(* IEC 61131-3 sources: daoli-st-library/DL_Process (part 28) *)

(* ---- FB_DL_ChillerYearWinStart.st ---- *)
(*==============================================================================
 * 组件名称 (Component)  : FB_DL_ChillerYearWinStart
 * 所属子库 (Sublibrary) : DL_Process
 * 当前版本 (Version)    : 1.0.0
 * 兼容性 (Platform)     : CODESYS 3.5+ / TwinCAT 3 / 汇川 InoProShop / 施耐德 Machine Expert
 *                         仅依赖 Standard.library（R_TRIG），零厂商私有库
 * 功能描述 (Function)   : 冷机年度启停窗与保养互锁。启动申请仅在「年窗电平
 *                         内 + 保养完成互锁成立」时放行 bRun，否则拒绝并按
 *                         独立成因（非窗 / 保养未完）给出 bBlocked 电平与
 *                         eBlock 成因（R190 归因唯一）；运行中可随时停止。
 *                         与 YearWindowCheck（年窗原子）分工：本件叠加
 *                         「非窗禁启」的设备控制语义。
 * 来源标签 (Origin)     : ROADMAP §16.5 R11 池（L725），自研 clean-room
 * 边界语义 (Boundary)   : ① 启动判据全组合闸（窗电平 / 保养互锁 / 无故障），
 *                         拒启不锁存故障（拒绝是正常业务态）；
 *                         ② 保养互锁输入非有限无涉（布尔域），无浮点量；
 *                         ③ eBlock 成因独立成员逐拍重算（拒绝成因随当前
 *                         条件实时回放，信息级允许每拍重算，R189）。
 * 输出语义 (Fallback)   : 【R191】bEnable = FALSE → bRun 强制 FALSE（启停
 *                         出口失能必须收敛）；eFault 相 → bRun FALSE + bError。
 * 码位     (Codes)      : 按 R297 范式零 16# 码位硬编码；错误出口 BOOL+ENUM(eCause)。
 * 红线自检 (Redline)    : 7 项红线已自检：R1 零全局 ✓｜R2 零物理地址 ✓｜R3 纯 IEC ✓
 *                         R4 无浮点域/组态无涉 ✓｜R5 双语同行注释 ✓
 *                         R6 CASE 带 ELSE 兜底迁 eFault ✓｜R7 R_TRIG 段 0 无条件刷新 ✓
 * 验收向量 (Acceptance) : V1 窗内 + 保养完 + 申请沿 → bRun=TRUE，bBlocked=FALSE；
 *                         V2 窗外申请沿 → bRun=FALSE，bBlocked=TRUE，
 *                         eBlock=eNotInWin；
 *                         V3 窗内但保养未完 → eBlock=eMaintDue（非窗成因
 *                         不再误报）。
 * 修订历史 (Revision)   : 2026-11-20  v1.0.0  R51 首版（批 2 · 序号 7）
 *==============================================================================*)
TYPE E_DL_CwsBlock :
(
    eNone     := 0,                          (* 无拒绝（已放行或无申请） / No block *)
    eNotInWin := 1,                          (* 非年窗禁启 / Not in year window *)
    eMaintDue := 2                           (* 保养未完禁启 / Maintenance interlock open *)
);
END_TYPE

TYPE E_DL_CwsState :
(
    eIdle  := 0,                             (* 停机待窗 / Idle *)
    eRun   := 10,                            (* 运行 / Running *)
    eFault := 90                             (* 故障锁存相 / Fault latched phase *)
);
END_TYPE

TYPE E_DL_CwsCause :
(
    eNone     := 0,                          (* 无故障成因 / No cause *)
    ePhaseBad := 3                           (* 非法相位兜底 / Illegal phase fallback *)
);
END_TYPE

FUNCTION_BLOCK FB_DL_ChillerYearWinStart
VAR_INPUT
    bInWin     : BOOL := FALSE;              (* 年窗电平（上层 YearWindowCheck 供给）[-] / Year-window level *)
    bMaintOk   : BOOL := TRUE;               (* 保养完成互锁电平 [-] / Maintenance interlock *)
    bStartReq  : BOOL := FALSE;              (* 启动申请电平 [-] / Start request *)
    bStopReq   : BOOL := FALSE;              (* 停止申请电平（运行中随时可停）[-] / Stop request *)
    bEnable    : BOOL := TRUE;               (* 使能 [-] / Enable *)
    bReset     : BOOL := FALSE;              (* 复位命令，上升沿清全部 [-] / Reset command *)
END_VAR
VAR_OUTPUT
    bRun       : BOOL;                       (* 冷机运行出口 [-] / Run outlet *)
    bStartOk   : BOOL;                       (* 本次申请放行单拍位 [-] / Start-allowed pulse *)
    bBlocked   : BOOL;                       (* 申请被拒电平（申请期实时）[-] / Blocked level *)
    eBlock     : E_DL_CwsBlock;              (* 拒绝成因（信息级逐拍重算，R189） / Block cause *)
    nRunCycles : UDINT;                      (* 累计启动次数 [次] / Run cycle count *)
    eState     : E_DL_CwsState;              (* 状态出口 / State outlet *)
    eCause     : E_DL_CwsCause;              (* 故障成因出口 / Fault cause outlet *)
    bError     : BOOL;                       (* 故障锁存标志 [-] / Fault latch flag *)
END_VAR
VAR
    _eState   : E_DL_CwsState := E_DL_CwsState.eIdle;     (* 内部相位（CASE 唯一写入目标） / Internal phase *)
    _eCause   : E_DL_CwsCause := E_DL_CwsCause.eNone;     (* 故障成因锁存量 / Latched cause *)
    rtStart   : R_TRIG;                      (* 启动申请沿实例，段 0 无条件调用 / Start edge instance *)
    rtStop    : R_TRIG;                      (* 停止申请沿实例，段 0 无条件调用 / Stop edge instance *)
    rtReset   : R_TRIG;                      (* 复位沿实例，段 0 无条件调用 / Reset edge instance *)
    _nCycles  : UDINT;                       (* 启动计数锁存 [次] / Cycle count latch *)
    _bStartOk : BOOL;                        (* 放行单拍量 [-] / Start-allowed work *)
    _bFault   : BOOL;                        (* 故障锁存位 / Latched fault bit *)
END_VAR

(* —— 段 0：沿实例无条件刷新（R228A；纯布尔域无浮点组态闸） —— *)
rtStart(CLK := bStartReq);                   (* 启动沿每拍必调 / Start edge every scan *)
rtStop(CLK := bStopReq);                     (* 停止沿每拍必调 / Stop edge every scan *)
rtReset(CLK := bReset);                      (* 复位沿每拍必调 / Reset edge every scan *)

(* —— 段 1：单拍量预清零（R107） —— *)
_bStartOk := FALSE;                          (* 放行脉冲预清，唯一分支置位 / Start-ok preset *)
bStartOk := FALSE;                           (* 放行出口预清 / Start-ok outlet preset *)
bBlocked := FALSE;                           (* 拒绝电平预清 / Blocked preset *)
eBlock := E_DL_CwsBlock.eNone;               (* 拒绝成因预清（判定分支覆盖） / Block cause preset *)

(* —— 段 2：复位沿处理（作用域：清故障 + 清计数 + 迁 eIdle（bRun 随相位收敛），R283 逐项声明） —— *)
IF rtReset.Q THEN
    _bFault := FALSE;                        (* 清故障锁存 / Clear fault *)
    _eCause := E_DL_CwsCause.eNone;          (* 清成因 / Clear cause *)
    _nCycles := 0;                           (* 清启动计数 / Clear count *)
    _eState := E_DL_CwsState.eIdle;          (* 迁停机相 / Back to idle *)
END_IF

(* —— 段 4：CASE 主状态机（ELSE 兜底迁 eFault，红线 6） —— *)
CASE _eState OF
    E_DL_CwsState.eIdle:                     (* 停机相 / Idle *)
        IF rtStart.Q AND bEnable THEN        (* 申请沿：判组合闸 / On start edge *)
            IF NOT bInWin THEN
                bBlocked := TRUE;            (* 拒绝电平 / Blocked level *)
                eBlock := E_DL_CwsBlock.eNotInWin;   (* 成因：非窗（独立成员，R190） / Cause: not in window *)
            ELSIF NOT bMaintOk THEN
                bBlocked := TRUE;            (* 拒绝电平 / Blocked level *)
                eBlock := E_DL_CwsBlock.eMaintDue;   (* 成因：保养未完 / Cause: maintenance *)
            ELSE
                _bStartOk := TRUE;           (* 放行单拍 / Start-ok pulse *)
                _nCycles := _nCycles + 1;    (* 启动计数（UDINT 回绕工程安全） / Count start *)
                _eState := E_DL_CwsState.eRun;   (* 进入运行 / Enter run *)
            END_IF
        END_IF
    E_DL_CwsState.eRun:                      (* 运行相：停止沿随时出 / Run *)
        IF rtStop.Q OR (NOT bEnable) THEN    (* 停止沿或失能：回停机 / Stop or disable *)
            _eState := E_DL_CwsState.eIdle;  (* 回停机相 / Back to idle *)
        END_IF
    E_DL_CwsState.eFault:                    (* 故障相：仅复位沿出（bRun 随段 5 收敛） / Fault *)
        ;                                    (* 锁存回放（R28） / Replay from latch *)
    ELSE                                     (* 非法相位兜底迁安全态 / Illegal phase fallback *)
        _eState := E_DL_CwsState.eFault;     (* 迁故障相 / To fault *)
        _bFault := TRUE;                     (* 同步锁存 / Latch *)
        _eCause := E_DL_CwsCause.ePhaseBad;  (* 成因：非法相位 / Cause: illegal phase *)
END_CASE

(* —— 段 5：出口映射（bRun 与相位同源同义，R191 名实双出口） —— *)
bRun := (_eState = E_DL_CwsState.eRun) AND bEnable AND (NOT _bFault);   (* 运行出口（失能/故障收敛 FALSE） / Run outlet *)
bStartOk := _bStartOk;                       (* 放行脉冲出口 / Start-ok outlet *)
nRunCycles := _nCycles;                      (* 启动计数出口 / Count outlet *)
bError := _bFault;                           (* 故障标志镜像 / Fault flag mirror *)
eState := _eState;                           (* 状态出口 / State outlet *)
eCause := _eCause;                           (* 成因出口 / Cause outlet *)
END_FUNCTION_BLOCK

(* ---- FB_DL_CleanRoomPressure.st ---- *)
(*==============================================================================
 * 组件名称 (Component)  : FB_DL_CleanRoomPressure
 * 所属子库 (Sublibrary) : DL_Process
 * 前缀     (Prefix)     : FB_DL_
 * 当前版本 (Version)    : 1.0.0
 * 兼容性   (Platform)   : CODESYS 3.5 / TwinCAT 3 / 汇川 InoProShop / Schneider
 *                         Machine Expert；纯 IEC 61131-3（第 3 版），
 *                         仅依赖标准库 MAX / MIN，零厂商方言、零定时器依赖
 * 作者     (Author)     : 道莅代码库 · PLC编程专家（R31）
 * 开源溯源 (Origin)     : 洁净室压差梯级控制公开工艺语义（行业池），道莅
 *                         clean-room 防御性实现，未复制任何外部源码行
 * 功能描述 (Function)   : 多房间正压梯级控制防倒流件。梯度校验先于控制：
 *                         逐室核对设定梯度沿洁净度递减方向严格递减，
 *                         倒置即锁存倒置标志并冻结投切（防倒流最高优先）；
 *                         控制层各室独立带回差双限：低于下限请求加大风量、
 *                         高于上限撤回请求、带内保持。
 * 码位     (Codes)      : 16#0005_00A3 信息级：压差/设定非有限该室退出仲裁、
 *                                      房间计数钳位（不置 bError）
 *                         16#0005_00A4 故障级：梯度倒置（锁存，独立复位通道）
 *                         16#0005_00A5~00A7 保留未启用（码表与实现对齐）
 * 边界防错 (Boundary)   : 1 梯度倒置锁存有可达解除式：独立 bRstInv 复位沿，
 *                           复位通道不受 NOT bEn 屏蔽（终审两式之一）；
 *                         2 房间计数钳上限、越界逐位清零；
 *                         3 非有限压差该室退出仲裁保持原投切并计掩码；
 *                         4 首拍全 FALSE；
 *                         5 无定时器/边沿实例（纯组合投切层）。
 * 修订历史 (Revision)   : 2026-11-18 v1.0.0 首版入库（R31 · 阶段三 · 序 13）
 *==============================================================================*)

(*==============================================================================
 * 功能块: FB_DL_CleanRoomPressure
 * 调用约定: 每个扫描周期无条件调用一次；压差与梯度设定经引脚数组注入，
 *           数组维度 1..8（8 室上限），有效室数经 uRoomCnt 给出。
 *==============================================================================*)
FUNCTION_BLOCK FB_DL_CleanRoomPressure
VAR_INPUT
    afDp    : ARRAY[1..8] OF REAL;    // 各室实测压差 [帕] / Per-room measured differential pressure [Pa]
    afSet   : ARRAY[1..8] OF REAL;    // 各室压差梯度设定 [帕]，须严格递减 / Per-room gradient setpoints [Pa], strictly decreasing
    uRoomCnt: UINT := 8;              // 有效房间数 [间]，合法域 1..8 / Valid room count, valid 1..8
    fBand   : REAL := 5.0;            // 回差半带宽 [帕] / Hysteresis half band [Pa]
    bEn     : BOOL := FALSE;          // 使能 / Enable flag
    bRstInv : BOOL := FALSE;          // 梯度倒置独立复位沿（不受使能屏蔽）/ Inversion reset edge, never masked by enable
END_VAR
VAR_OUTPUT
    abBoost : ARRAY[1..8] OF BOOL;    // 各室加大风量请求 / Per-room boost request
    bInvert : BOOL;                   // 梯度倒置锁存标志 / Gradient inversion latch flag
    uErrorId: UDINT;                  // 错误码，0 = 无错 / Error code, 0 = none
END_VAR
VAR
    rTrigRst: R_TRIG;                 // 倒置复位沿检测，每拍无条件刷新 / Inversion reset edge detector
    uCntEff : INT;                    // 钳位后有效室数 [间]，INT 域循环 / Effective clamped room count, INT domain
    i       : INT;                    // 逐室循环索引 / Per-room loop index
    bRoomOk : ARRAY[1..8] OF BOOL;    // 各室数据有效掩码 / Per-room data validity mask
    bBadAny : BOOL;                   // 任一室数据无效 / Any room data invalid
    bFirst  : BOOL := TRUE;           // 首拍标志 / First-scan flag
    fLo     : REAL;                   // 本室投切下限 [帕] / Room switching lower bound [Pa]
    fHi     : REAL;                   // 本室投切上限 [帕] / Room switching upper bound [Pa]
END_VAR
VAR CONSTANT
    DL_CRP_ROOM_MAX: INT  := 8;       // 房间数上限 [间] / Room count upper bound
    DL_CRP_FIN     : REAL := 1.0E30;  // REAL 有限幅值判界 / REAL finiteness magnitude bound
END_VAR

// ---- 段 1｜边沿实例无条件刷新（红线：禁入条件分支）----------------------------
rTrigRst(CLK := bRstInv);                             // 倒置复位沿检测 / Inversion reset edge detection

// ---- 段 2｜梯度倒置独立复位：先于一切使能门控（R38 复位通道不屏蔽）--------------
IF rTrigRst.Q THEN
    bInvert := FALSE;                                 // 复位清倒置锁存 / Reset clears inversion latch
END_IF

// ---- 段 3｜计数钳位与首拍初始化 --------------------------------------------------
uCntEff := MIN(UINT_TO_INT(uRoomCnt), DL_CRP_ROOM_MAX); // 计数钳上限，统一 INT 域 / Clamp count, unified INT domain
uCntEff := MAX(uCntEff, 1);                           // 下限保 1 防 0 循环 / Floor at 1 against empty loop
IF bFirst THEN
    FOR i := 1 TO DL_CRP_ROOM_MAX DO
        abBoost[i] := FALSE;                          // 首拍全 FALSE / First scan all FALSE
        bRoomOk[i] := TRUE;                           // 掩码预置有效 / Mask preset valid
    END_FOR
    bFirst := FALSE;                                  // 清首拍标志 / Clear first-scan flag
END_IF

// ---- 段 4｜梯度校验先于控制（防倒流最高优先）--------------------------------------
IF NOT bInvert THEN
    FOR i := 1 TO (uCntEff - 1) DO
        IF (afSet[i] <> afSet[i]) OR (afSet[i + 1] <> afSet[i + 1])
           OR (ABS(afSet[i]) >= DL_CRP_FIN) OR (ABS(afSet[i + 1]) >= DL_CRP_FIN) THEN
            bInvert := TRUE;                          // 非有限设定按倒置保守处理（留档）/ Non-finite set treated as inversion
        ELSIF afSet[i] <= afSet[i + 1] THEN
            bInvert := TRUE;                          // 梯度未严格递减判倒置 / Non-decreasing gradient is inversion
        END_IF
    END_FOR
END_IF

// ---- 段 5｜数据有效性掩码（非有限该室退出仲裁）------------------------------------
bBadAny := FALSE;                                     // 掩码标志先清 / Clear mask flag
FOR i := 1 TO DL_CRP_ROOM_MAX DO
    IF i <= uCntEff THEN
        bRoomOk[i] := (afDp[i] = afDp[i]) AND (ABS(afDp[i]) < DL_CRP_FIN); // 本室压差有限 / Room pressure finite
        bRoomOk[i] := bRoomOk[i] AND (fBand >= 0.0) AND (fBand < DL_CRP_FIN); // 带宽合法性并入 / Band legality merged
    ELSE
        bRoomOk[i] := FALSE;                          // 越界室退出并视为无效 / Out-of-range room excluded
        abBoost[i] := FALSE;                          // 越界逐位清零（R29 输出确定值）/ Out-of-range bits cleared
    END_IF
    IF (NOT bRoomOk[i]) AND (i <= uCntEff) THEN
        bBadAny := TRUE;                              // 有效域内存在无效室 / Invalid room inside valid range
    END_IF
END_FOR

// ---- 段 6｜控制层：各室独立带回差双限（倒置锁存期冻结投切保持原值）----------------
IF (NOT bInvert) AND bEn THEN
    FOR i := 1 TO uCntEff DO
        fLo := afSet[i] - fBand;                      // 本室下限 / Room lower bound
        fHi := afSet[i] + fBand;                      // 本室上限 / Room upper bound
        IF NOT bRoomOk[i] THEN
            abBoost[i] := abBoost[i];                 // 无效室退出仲裁保持原值 / Invalid room holds state
        ELSIF afDp[i] < fLo THEN
            abBoost[i] := TRUE;                       // 低于下限请求加大风量 / Below lower bound, boost on
        ELSIF afDp[i] > fHi THEN
            abBoost[i] := FALSE;                      // 高于上限撤回请求 / Above upper bound, boost off
        ELSE
            abBoost[i] := abBoost[i];                 // 带内保持（回差防抖）/ In band, hold
        END_IF
    END_FOR
END_IF

// ---- 段 7｜错误码装配：倒置锁存故障级优先，信息级居次 ------------------------------
IF bInvert THEN
    uErrorId := 16#0005_00A4;                         // 故障级：梯度倒置锁存 / Fault: inversion latched
ELSIF bBadAny OR (UINT_TO_INT(uRoomCnt) > DL_CRP_ROOM_MAX) THEN
    uErrorId := 16#0005_00A3;                         // 信息级：非有限/计数钳位 / Info: non-finite or count clamp
ELSE
    uErrorId := 16#0000_0000;                         // 无码 / No code
END_IF
END_FUNCTION_BLOCK

(* ---- FB_DL_CoagDoseJarTestSeq.st ---- *)
(*
  道莅工业代码库 / Daoli Industrial ST Library
  组件: FB_DL_CoagDoseJarTestSeq
  分类: DL_Process
  复杂度: C4 ｜ 版本: 1.0.0 ｜ 2026-11-24
  平台兼容: CODESYS 3.5+ / TwinCAT 3 / 汇川 InoProShop / 施耐德 Machine Expert
  开源溯源: 无（clean-room 工程公式自研；参考公开的混凝烧杯试验与投加量换算工艺公式，
            未复制任何受版权保护代码）
  许可证: 本项目自有 (MIT)

  功能职责:
    水厂混凝加药闭环。前馈按进水浊度三段给投加基准，烧杯试验结果到达后修正基准，
    沉后浊度复核超限则再整定（单次限幅 ±20%，最多 3 轮）。
    相序: eIdle →（bEnable 上升沿）eFeedForward → eJarTestWait → eTrim → eVerify
          →（达标 / 轮次耗尽）eHold；eJarTestWait 超时 → eFault（码 11）。

  输入/输出契约:
    IN  bEnable 上升沿启动；FALSE 撤销执行位 bDoseOn 并回 eIdle（设定值保留，见 R191 声明）。
    IN  bReset  上升沿是 eFault 的唯一出口（还须残留故障条件消失）。
    OUT rDoseLh 投加量设定 [L/h]，故障相与保持相输出「最后有效投加」而不掉零。
    OUT bDoseOn 投加执行位，故障相与 eHold 之外的活动相为 TRUE。

  码表 (Codes):
    11 = 烧杯结果等待超时（故障级；执行位 FALSE，但投加设定保持最后有效值不掉零）
    12 = 复核整定轮次耗尽（告警级；转 eHold 保持最后有效投加，不置故障相）
    13 = 烧杯结果非法（信息级；本拍跳过修正，基准不变）
    14 = 进水流量无效（故障级，rFlowM3h ≤ 0，投加量无法换算）
    15 = 母液浓度无效（故障级，rStockGL ≤ 0，除零闸拦截）
    16 = 沉后浊度设定无效（故障级，rOutNtuSp ≤ 0，复核倍率不可信）
    17 = 投加上限无效（故障级，rDoseMaxLh ≤ 0，无饱和载体）
    99 = 非法状态枚举值（ELSE 兜底）

  边界与红线:
    ① 两个 TON（tonJar / tonSettle）与三个 R_TRIG 全部在 CASE 外无条件刷新（R7），CASE 内只读 .Q。
    ② 两个 TON 的 IN 各自串本相闸（eJarTestWait / eVerify）并带 NOT .Q 自复位（R188），
       属「本相单发计时」而非跨相累计看门狗（红线 14 声明）。
    ③ R528：eIdle 只在 bEnable 上升沿且母液浓度/流量/投加上限三项均有效时才迁 eFeedForward；
       全默认引脚（全 0）时停留 eIdle，绝不直达前馈或投加相。
    ④ eFault 出口 = rtReset.Q AND NOT _bFaultCondNow（残留条件按锁存码逐条反算，R28 可达性）。
    ⑤ 单一状态机内联实现：无方法级封装、无属性段、无倒序循环、无数组透传
  修订历史: 2026-11-24  v1.0.0  R82-B 首版
*)

TYPE E_DL_COAG_STATE :
(
    eIdle        := 0,    // 空闲：等使能上升沿 / Idle: waiting for the enable rising edge
    eFeedForward := 1,    // 前馈相：按进水浊度三段给基准 / Feed-forward: base dose from three inlet turbidity bands
    eJarTestWait := 2,    // 烧杯等待相：等结果沿，超时转故障 / Jar test wait: waiting for the result edge, timeout goes to fault
    eTrim        := 3,    // 修正相：按烧杯结果单次限幅修正基准 / Trim: bounded correction of the base by the jar test result
    eVerify      := 4,    // 复核相：沉后浊度与设定比较 / Verify: compare the settled turbidity with the setpoint
    eHold        := 5,    // 保持相：保持最后有效投加等复位 / Hold: keep the last valid dose until reset
    eFault       := 6     // 故障安全相：执行位撤销，设定保持 / Fault safe phase: run bit withdrawn, setpoint kept
);
END_TYPE

FUNCTION_BLOCK FB_DL_CoagDoseJarTestSeq
VAR_INPUT
    bEnable         : BOOL := FALSE;      // 使能（上升沿启动；FALSE 撤销执行位回空闲）/ Enable, rising edge starts, FALSE withdraws the run bit
    bReset          : BOOL := FALSE;      // 复位（上升沿，eFault 唯一出口）/ Reset rising edge, the only fault exit
    bJarResultReady : BOOL := FALSE;      // 烧杯结果到达（上升沿有效）/ Jar test result ready, rising edge only
    rJarResultMgL   : REAL := 0.0;        // 烧杯试验最优投加浓度 [mg/L] / Jar test optimum dose concentration [mg/L]
    rInNtu          : REAL := 0.0;        // 进水浊度 [NTU] / Inlet turbidity [NTU]
    rOutNtu         : REAL := 0.0;        // 沉后浊度实测 [NTU] / Settled outlet turbidity [NTU]
    rOutNtuSp       : REAL := 0.0;        // 沉后浊度设定 [NTU] / Settled turbidity setpoint [NTU]
    rFlowM3h        : REAL := 0.0;        // 进水流量 [m3/h] / Inlet flow [m3/h]
    rStockGL        : REAL := 0.0;        // 母液浓度 [g/L]（1 g/L = 1 kg/m3）/ Stock concentration [g/L]
    rDoseMaxLh      : REAL := 0.0;        // 投加泵上限 [L/h] / Dosing pump upper limit [L/h]
    tSettleTime     : TIME := T#15M;      // 沉后稳定等待，有效域 100ms..2h [s] / Settling wait, valid domain 100ms..2h
    tVerifyTimeout  : TIME := T#30M;      // 烧杯结果等待超时，有效域 100ms..2h [s] / Jar result timeout, valid domain 100ms..2h
END_VAR
VAR_OUTPUT
    rDoseLh         : REAL := 0.0;        // 投加量设定 [L/h] / Dose setpoint [L/h]
    bDoseOn         : BOOL := FALSE;      // 投加执行位（故障相强制 FALSE）/ Dose run bit, forced FALSE in the fault phase
    iErrCode        : INT := 0;           // 错误码（故障期锁存回放，非故障期为信息码）/ Error code, latched replay during fault
    sMsg            : STRING;             // 文本提示（当前相位摘要）/ Text message, a summary of the current phase
END_VAR
VAR
    _eState         : E_DL_COAG_STATE := E_DL_COAG_STATE.eIdle;   // 内部相位（CASE 唯一写入目标）/ Internal phase, the only CASE write target
    _bFaultLatch    : BOOL := FALSE;      // 故障锁存位（仅复位出口清除）/ Fault latch, cleared only at the reset exit
    _iErrLatch      : INT := 0;           // 锁存故障码（故障期唯一回放源）/ Latched fault code, the only replay source during fault
    _iInfoCode      : INT := 0;           // 信息级/告警级码（永不进故障锁存）/ Info or warning code, never latched as a fault
    _iErrTmp        : INT := 0;           // 当拍故障首因中间量 / First fault cause of this scan
    _bFaultReq      : BOOL := FALSE;      // 当拍故障请求（段 7 统一锁存）/ Fault request of this scan, latched at segment 7
    _bFaultCondNow  : BOOL := FALSE;      // 残留故障条件（eFault 出口唯一附加判据）/ Residual fault condition, the only extra fault-exit criterion
    _rBaseMgL       : REAL := 0.0;        // 当前投加基准浓度 [mg/L] / Current base dose concentration [mg/L]
    _rDoseCmd       : REAL := 0.0;        // 当拍换算投加量 [L/h] / Dose computed this scan [L/h]
    _rDoseLastGood  : REAL := 0.0;        // 最后有效投加量 [L/h]（不掉零载体）/ Last valid dose [L/h], the never-zero carrier
    _rInNtuCl       : REAL := 0.0;        // 进水浊度净化副本 [NTU] / Sanitised inlet turbidity copy [NTU]
    _rOutNtuCl      : REAL := 0.0;        // 沉后浊度净化副本 [NTU] / Sanitised settled turbidity copy [NTU]
    _rDelta         : REAL := 0.0;        // 基准修正相对偏差（无量纲）/ Relative correction of the base, dimensionless
    _rRatio         : REAL := 0.0;        // 浊度复核倍率（无量纲）/ Turbidity verification ratio, dimensionless
    _iTrimCnt       : INT := 0;           // 整定轮次计数，容量载体 DL_CDJ_CYCLE_MAX [次] / Trim round counter, capacity carrier DL_CDJ_CYCLE_MAX [count]
    _tSettle        : TIME := T#15M;      // 沉后稳定等待钳定值 [s] / Clamped settling wait [s]
    _tVerify        : TIME := T#30M;      // 烧杯超时钳定值 [s] / Clamped jar timeout [s]
    rtReset         : R_TRIG;             // bReset 边沿（段 3 无条件刷新）/ bReset edge, refreshed unconditionally at segment 3
    rtEnable        : R_TRIG;             // bEnable 边沿（段 3 无条件刷新）/ bEnable edge, refreshed unconditionally at segment 3
    rtJar           : R_TRIG;             // 烧杯结果边沿（段 3 无条件刷新）/ Jar result edge, refreshed unconditionally at segment 3
    tonJar          : TON;                // 烧杯等待计时（本相单发，自复位）/ Jar wait timer, single shot in its phase with self reset
    tonSettle       : TON;                // 沉后稳定计时（本相单发，自复位）/ Settling timer, single shot in its phase with self reset
END_VAR
VAR CONSTANT
    DL_CDJ_EPS         : REAL := 1.0E-6;      // 除零闸阈值 [-] / Divide-by-zero guard threshold [-]
    DL_CDJ_FIN         : REAL := 1.0E15;      // 非有限判据阈值（ABS 比较用）[-] / Non-finite criterion threshold, compared by ABS [-]
    DL_CDJ_NTU_SPLIT1  : REAL := 20.0;        // 进水浊度第一分段阈值 [NTU] / First inlet turbidity band threshold [NTU]
    DL_CDJ_NTU_SPLIT2  : REAL := 50.0;        // 进水浊度第二分段阈值 [NTU] / Second inlet turbidity band threshold [NTU]
    DL_CDJ_MGL_LOW     : REAL := 8.0;         // 低浊段基准投加浓度 [mg/L] / Base dose concentration of the low band [mg/L]
    DL_CDJ_MGL_MID     : REAL := 15.0;        // 中浊段基准投加浓度 [mg/L] / Base dose concentration of the mid band [mg/L]
    DL_CDJ_MGL_HIGH    : REAL := 25.0;        // 高浊段基准投加浓度 [mg/L] / Base dose concentration of the high band [mg/L]
    DL_CDJ_TRIM_LIM    : REAL := 0.2;         // 单次修正限幅 ±20%（无量纲）/ Per-round correction limit of plus or minus twenty percent, dimensionless
    DL_CDJ_NTU_RATIO   : REAL := 1.15;        // 复核超限倍率（无量纲）/ Verification exceed factor, dimensionless
    DL_CDJ_CYCLE_MAX   : INT := 3;            // 整定轮次上限 [次] / Trim round upper limit [count]
    DL_CDJ_ONE         : INT := 1;            // 计数步进一 [1] / Counter step of one [1]
    DL_CDJ_ZERO        : INT := 0;            // 计数零基准 [-] / Counter zero base [-]
    DL_CDJ_T_MIN       : TIME := T#100MS;     // 时间参数下限 [s] / Time parameter lower bound [s]
    DL_CDJ_T_MAX       : TIME := T#2H;        // 时间参数上限 [s] / Time parameter upper bound [s]
    DL_CDJ_T_SETTLE_DEF: TIME := T#15M;       // 沉后等待默认回退值（本身在域内）[s] / Default settling wait, already inside the domain [s]
    DL_CDJ_T_VERIFY_DEF: TIME := T#30M;       // 烧杯超时默认回退值（本身在域内）[s] / Default jar timeout, already inside the domain [s]
END_VAR

(* —— 段 1：中间量预置（只清当拍扫描量，不清锁存/基准/最后有效投加，FB32-1） —— *)
_iErrTmp   := 0;                              // 当拍故障首因复位 / Scan first fault cause reset
_bFaultReq := FALSE;                          // 当拍故障请求复位 / Scan fault request reset

(* —— 段 2：时间参数两级回退 + 入参非有限兜底 + 残留故障条件反算 —— *)
IF (tSettleTime < DL_CDJ_T_MIN) OR (tSettleTime > DL_CDJ_T_MAX) THEN
    _tSettle := DL_CDJ_T_SETTLE_DEF;          // 越域：回一级默认常量 / Out of domain: fall back to the default constant
ELSE
    _tSettle := tSettleTime;                  // 域内：原值采用 / Inside the domain: use as given
END_IF
IF (tVerifyTimeout < DL_CDJ_T_MIN) OR (tVerifyTimeout > DL_CDJ_T_MAX) THEN
    _tVerify := DL_CDJ_T_VERIFY_DEF;          // 越域：回一级默认常量 / Out of domain: fall back to the default constant
ELSE
    _tVerify := tVerifyTimeout;               // 域内：原值采用 / Inside the domain: use as given
END_IF
_rInNtuCl := rInNtu;                          // 进水浊度副本，参与前馈分段 / Inlet turbidity copy used by the feed-forward bands
IF (ABS(_rInNtuCl) > DL_CDJ_FIN) OR (_rInNtuCl < 0.0) THEN
    _rInNtuCl := 0.0;                         // 非有限或负值兜底为零（非有限判据用 ABS>FIN）/ Non-finite or negative falls back to zero
END_IF
_rOutNtuCl := rOutNtu;                        // 沉后浊度副本，参与复核倍率 / Settled turbidity copy used by the verification ratio
IF (ABS(_rOutNtuCl) > DL_CDJ_FIN) OR (_rOutNtuCl < 0.0) THEN
    _rOutNtuCl := 0.0;                        // 非有限或负值兜底为零 / Non-finite or negative falls back to zero
END_IF
_bFaultCondNow := FALSE;                      // 残留条件预置（eFault 出口唯一附加判据）/ Residual preset, the only extra fault-exit criterion
IF _iErrLatch = 14 THEN
    _bFaultCondNow := (rFlowM3h <= 0.0);      // 码 14：流量仍未恢复 / Code 14: flow still invalid
ELSIF _iErrLatch = 15 THEN
    _bFaultCondNow := (rStockGL <= DL_CDJ_EPS);      // 码 15：浓度仍未恢复 / Code 15: concentration still invalid
ELSIF _iErrLatch = 16 THEN
    _bFaultCondNow := (ABS(rOutNtuSp) <= DL_CDJ_EPS);  // 码 16：设定仍未恢复 / Code 16: setpoint still invalid
ELSIF _iErrLatch = 17 THEN
    _bFaultCondNow := (rDoseMaxLh <= DL_CDJ_EPS);    // 码 17：上限仍未恢复 / Code 17: upper limit still invalid
END_IF
(* 码 11（等待超时）是一次性已消费事件、码 99 是内部枚举损坏，二者均无残留输入条件，
   故复位沿单独即可退出故障相；此两条可达路径在上表已显式穷举，无死锁。 / Codes 11 and 99 leave no residual input condition *)

(* —— 段 3：边沿与定时器（全部在 CASE 外无条件刷新，R7；IN 带 NOT .Q 自复位，R188） —— *)
rtReset(CLK := bReset);                       // 复位边沿无条件刷新 / Reset edge refreshed unconditionally
rtEnable(CLK := bEnable);                     // 使能边沿无条件刷新（R528 起点判据）/ Enable edge refreshed unconditionally
rtJar(CLK := bJarResultReady);                // 烧杯结果边沿无条件刷新 / Jar result edge refreshed unconditionally
tonJar(IN := (_eState = E_DL_COAG_STATE.eJarTestWait) AND (NOT tonJar.Q) AND (NOT _bFaultLatch),
       PT := _tVerify);                       // 本相单发计时：仅等待相计时，超时即迁故障 / Single-shot timer in the wait phase only
tonSettle(IN := (_eState = E_DL_COAG_STATE.eVerify) AND (NOT tonSettle.Q) AND (NOT _bFaultLatch),
          PT := _tSettle);                    // 本相单发计时：仅复核相计时，与等待相无关 / Single-shot timer in the verify phase only

(* —— 段 4：状态机主体（唯一相位写入点；故障只置请求，锁存与迁相由段 7 执行） —— *)
CASE _eState OF
    E_DL_COAG_STATE.eIdle :
        (* 迁移①：拍 N 进入（使能上升沿）/ 本拍行为：三项参数有效性校验，任一无效即进故障 / 拍 N+1 转出至前馈相 *)
        IF rtEnable.Q AND (NOT _bFaultLatch) THEN
            IF rStockGL <= DL_CDJ_EPS THEN
                _iErrTmp   := 15;                                  // 故障级：母液浓度无效（除零闸）/ Fault: invalid stock concentration
                _bFaultReq := TRUE;                                 // 请求段 7 锁存 / Request the latch at segment 7
            ELSIF rFlowM3h <= 0.0 THEN
                _iErrTmp   := 14;                                  // 故障级：进水流量无效 / Fault: invalid inlet flow
                _bFaultReq := TRUE;                                 // 请求段 7 锁存 / Request the latch at segment 7
            ELSIF rDoseMaxLh <= DL_CDJ_EPS THEN
                _iErrTmp   := 17;                                  // 故障级：投加上限无效 / Fault: invalid pump upper limit
                _bFaultReq := TRUE;                                 // 请求段 7 锁存 / Request the latch at segment 7
            ELSE
                _iTrimCnt  := DL_CDJ_ZERO;                          // 新周期：整定轮次归零 / New cycle: trim counter cleared
                _iInfoCode := 0;                                    // 新周期：信息码归零 / New cycle: info code cleared
                _eState    := E_DL_COAG_STATE.eFeedForward;         // 迁移①：进前馈相 / Move to feed-forward
            END_IF
        END_IF

    E_DL_COAG_STATE.eFeedForward :
        (* 迁移②：拍 N 进入 / 本拍行为：按进水浊度三段给投加基准 / 拍 N+1 转出至烧杯等待相 *)
        IF _rInNtuCl <= DL_CDJ_NTU_SPLIT1 THEN
            _rBaseMgL := DL_CDJ_MGL_LOW;                            // 低浊段基准 [mg/L] / Low band base [mg/L]
        ELSIF _rInNtuCl <= DL_CDJ_NTU_SPLIT2 THEN
            _rBaseMgL := DL_CDJ_MGL_MID;                            // 中浊段基准 [mg/L] / Mid band base [mg/L]
        ELSE
            _rBaseMgL := DL_CDJ_MGL_HIGH;                           // 高浊段基准 [mg/L] / High band base [mg/L]
        END_IF
        _eState := E_DL_COAG_STATE.eJarTestWait;                    // 迁移②：进等待相 / Move to the jar wait phase

    E_DL_COAG_STATE.eJarTestWait :
        (* 迁移③：本拍合法事件（结果沿）优先于超时（R275）/ 拍 N 进入 / 拍 N+1 转出至修正相或故障相 *)
        IF rtJar.Q THEN
            _eState := E_DL_COAG_STATE.eTrim;                       // 迁移③：进修正相 / Move to the trim phase
        ELSIF tonJar.Q THEN
            _iErrTmp   := 11;                                       // 故障级：等待超时（设定保持不掉零）/ Fault: wait timeout, the setpoint is kept
            _bFaultReq := TRUE;                                     // 请求段 7 锁存 / Request the latch at segment 7
        END_IF

    E_DL_COAG_STATE.eTrim :
        (* 迁移④：拍 N 进入 / 本拍行为：按烧杯结果单次限幅 ±20% 修正基准、轮次饱和计数 / 拍 N+1 转出至复核相 *)
        _iInfoCode := 0;                                            // 进入修正：信息码归零 / Entering trim: info code cleared
        IF _iTrimCnt < DL_CDJ_CYCLE_MAX THEN
            _iTrimCnt := _iTrimCnt + DL_CDJ_ONE;                    // 轮次净额 +1，达容量上限即饱和 / Net round increment, saturated at capacity
        END_IF
        // NaN 与任何数比较均为假，故用 NOT(正向域) 做兜底，NaN 必落进非法分支
        IF NOT ((rJarResultMgL > DL_CDJ_EPS) AND (rJarResultMgL <= DL_CDJ_FIN)) THEN
            _iInfoCode := 13;                                       // 信息级：结果非法，本拍不改基准 / Info: illegal result, the base is untouched
        ELSIF _rBaseMgL > DL_CDJ_EPS THEN
            // 量纲: (mg/L - mg/L)/(mg/L) = 无量纲相对偏差，乘基准得新基准 [mg/L]
            _rDelta := (rJarResultMgL - _rBaseMgL) / _rBaseMgL;      // 相对偏差（分母已闸）/ Relative deviation, the denominator is guarded
            IF ABS(_rDelta) > DL_CDJ_FIN THEN
                _rDelta := 0.0;                                      // 偏差非有限即弃用，保基准 / non-finite deviation discarded
            END_IF
            IF _rDelta > DL_CDJ_TRIM_LIM THEN
                _rDelta := DL_CDJ_TRIM_LIM;                         // 正向限幅 +20% / Positive clamp at plus twenty percent
            END_IF
            IF _rDelta < -(DL_CDJ_TRIM_LIM) THEN
                _rDelta := -(DL_CDJ_TRIM_LIM);                      // 负向限幅 -20% / Negative clamp at minus twenty percent
            END_IF
            _rBaseMgL := _rBaseMgL * (1.0 + _rDelta);               // 量纲: (mg/L)*(无量纲) = mg/L / (mg/L) times dimensionless gives mg/L
        END_IF
        _eState := E_DL_COAG_STATE.eVerify;                         // 迁移④：进复核相 / Move to the verify phase

    E_DL_COAG_STATE.eVerify :
        (* 迁移⑤⑥：拍 N 进入 / 本拍行为：稳定后比较沉后浊度与设定，超 1.15 倍回修正 / 拍 N+1 转出至修正或保持相 *)
        IF tonSettle.Q THEN
            IF ABS(rOutNtuSp) <= DL_CDJ_EPS THEN
                _iErrTmp   := 16;                                   // 故障级：设定无效，倍率不可信 / Fault: invalid setpoint, the ratio is untrustworthy
                _bFaultReq := TRUE;                                 // 请求段 7 锁存 / Request the latch at segment 7
            ELSE
                // 量纲: (NTU)/(NTU) = 无量纲倍率，与 1.15 无量纲阈值直比
                _rRatio := _rOutNtuCl / rOutNtuSp;                  // 复核倍率（分母已闸）/ Verification ratio with a guarded denominator
                IF _rRatio > DL_CDJ_NTU_RATIO THEN
                    IF _iTrimCnt >= DL_CDJ_CYCLE_MAX THEN
                        _iInfoCode := 12;                           // 告警级：轮次耗尽，转保持 / Warning: rounds exhausted, go to hold
                        _eState    := E_DL_COAG_STATE.eHold;        // 迁移⑥：保持最后有效投加 / Keep the last valid dose
                    ELSE
                        _eState := E_DL_COAG_STATE.eTrim;           // 迁移⑤：回修正相再整定 / Back to trim for another round
                    END_IF
                ELSE
                    _iInfoCode := 0;                                // 达标：清信息码 / Passed: info code cleared
                    _eState    := E_DL_COAG_STATE.eHold;            // 迁移⑤：达标转保持相 / Passed, go to hold
                END_IF
            END_IF
        END_IF

    E_DL_COAG_STATE.eHold :
        (* 迁移⑦：拍 N 进入（复核达标或轮次耗尽）/ 本拍行为：执行位保持、设定保持 / 拍 N+1 转出至 eIdle（复位沿） *)
        IF rtReset.Q THEN
            _iInfoCode := 0;                                        // 复位：清信息码 / Reset: info code cleared
            _eState    := E_DL_COAG_STATE.eIdle;                    // 迁移⑦：回空闲相，不滞留 / Back to idle, never parked
        END_IF

    E_DL_COAG_STATE.eFault :
        (* 迁移⑧：拍 N 进入 / 本拍行为：只等出口条件（复位沿 + 残留条件消失）/ 拍 N+1 转出至 eIdle *)
        IF rtReset.Q AND (NOT _bFaultCondNow) THEN
            _bFaultLatch := FALSE;                                  // 清故障锁存 / Clear the fault latch
            _iErrLatch   := 0;                                      // 清锁存故障码 / Clear the latched code
            _iInfoCode   := 0;                                      // 清信息码 / Clear the info code
            _iTrimCnt    := DL_CDJ_ZERO;                            // 整定轮次清零 / Trim counter cleared
            _eState      := E_DL_COAG_STATE.eIdle;                  // 回空闲相 / Back to idle
        END_IF
ELSE
    (* 迁移⑨：非法枚举兜底（R6），码位赋值与锁存 3 行内配对（R45） *)
    IF NOT _bFaultLatch THEN
        _iErrLatch   := 99;                                         // 故障级：非法状态枚举值 / Fault: illegal state enum value
        _bFaultLatch := TRUE;                                       // 置故障锁存 / Latch the fault
    END_IF
END_CASE

(* —— 段 5：投加量换算（CASE 之后单点重算，使本拍更新的基准立刻生效，FB33-1） —— *)
IF (rStockGL > DL_CDJ_EPS) AND (rFlowM3h > 0.0) THEN
    // 量纲: (mg/L)*(m3/h)/1000 = kg/h 干药剂；(kg/h) / (g/L = kg/m3) * 1000 L/m3 = L/h 母液
    _rDoseCmd := _rBaseMgL * rFlowM3h / rStockGL;                   // 投加体积流量 [L/h] / Dosing volume flow [L/h]
    IF _rDoseCmd > rDoseMaxLh THEN
        _rDoseCmd := rDoseMaxLh;                                    // 上限饱和（载体 rDoseMaxLh）/ Saturate at the pump limit
    END_IF
    IF _rDoseCmd < 0.0 THEN
        _rDoseCmd := 0.0;                                           // 下限饱和 / Saturate at zero
    END_IF
ELSE
    _rDoseCmd := 0.0;                                               // 分母或流量无效：出零不猜值 / Invalid denominator or flow: emit zero, never guess
END_IF

(* —— 段 6：最后有效投加跟踪（不掉零载体，仅活动相且命令为正值时刷新） —— *)
IF (NOT _bFaultLatch) AND (_rDoseCmd > 0.0) THEN
    IF (_eState = E_DL_COAG_STATE.eFeedForward) OR (_eState = E_DL_COAG_STATE.eJarTestWait)
       OR (_eState = E_DL_COAG_STATE.eTrim) OR (_eState = E_DL_COAG_STATE.eVerify) THEN
        _rDoseLastGood := _rDoseCmd;                                // 每次相迁移与在线运行均刷新 / Refreshed on every phase move and while running
    END_IF
END_IF

(* —— 段 7：故障锁存 + 段尾故障迁相 + 撤使能降级（R191：已声明为「降级 + 设定保留」） —— *)
IF _bFaultReq AND (NOT _bFaultLatch) THEN
    _iErrLatch   := _iErrTmp;                                       // 锁存当拍首因 / Latch the first cause of this scan
    _bFaultLatch := TRUE;                                           // 置故障锁存 / Latch the fault
END_IF
IF _bFaultLatch AND (_eState <> E_DL_COAG_STATE.eFault) THEN
    _eState := E_DL_COAG_STATE.eFault;                              // 锁存即迁相（段尾统一执行）/ The latch forces the fault phase at the tail
END_IF
IF (NOT bEnable) AND (NOT _bFaultLatch) AND (_eState <> E_DL_COAG_STATE.eIdle) THEN
    _eState := E_DL_COAG_STATE.eIdle;                               // 撤使能：回空闲，设定值保留 / Disable: back to idle with the setpoint kept
END_IF

(* —— 段 8：统一出口（单点映射，禁在 CASE 后无条件清零 CASE 内赋值标识符，FB33-1） —— *)
bDoseOn := (NOT _bFaultLatch) AND ((_eState = E_DL_COAG_STATE.eFeedForward)
           OR (_eState = E_DL_COAG_STATE.eJarTestWait) OR (_eState = E_DL_COAG_STATE.eTrim)
           OR (_eState = E_DL_COAG_STATE.eVerify) OR (_eState = E_DL_COAG_STATE.eHold));  // 执行位：故障相强制 FALSE / Run bit, forced FALSE in fault
IF _bFaultLatch OR (_eState = E_DL_COAG_STATE.eHold) THEN
    rDoseLh := _rDoseLastGood;                                      // 故障相与保持相：设定保持最后有效值不掉零 / Fault and hold keep the last valid setpoint
ELSE
    rDoseLh := _rDoseCmd;                                           // 活动相：输出当拍换算值 / Active phases emit the freshly computed dose
END_IF
IF _bFaultLatch THEN
    iErrCode := _iErrLatch;                                         // 故障期回放锁存码 / Replay the latched code during fault
ELSE
    iErrCode := _iInfoCode;                                         // 非故障期输出信息/告警码 / Info or warning code outside fault
END_IF
IF _eState = E_DL_COAG_STATE.eIdle THEN
    sMsg := 'IDLE';                                                 // 空闲 / Idle
ELSIF _eState = E_DL_COAG_STATE.eFeedForward THEN
    sMsg := 'FEEDFWD';                                              // 前馈给定 / Feed-forward
ELSIF _eState = E_DL_COAG_STATE.eJarTestWait THEN
    sMsg := 'JARWAIT';                                              // 等烧杯结果 / Waiting for the jar result
ELSIF _eState = E_DL_COAG_STATE.eTrim THEN
    sMsg := 'TRIM';                                                 // 基准修正 / Base trimming
ELSIF _eState = E_DL_COAG_STATE.eVerify THEN
    sMsg := 'VERIFY';                                               // 沉后复核 / Settled verification
ELSIF _eState = E_DL_COAG_STATE.eHold THEN
    sMsg := 'HOLD';                                                 // 保持 / Holding
ELSE
    sMsg := 'FAULT';                                                // 故障 / Fault
END_IF
END_FUNCTION_BLOCK

(* ---- FB_DL_CoaterGapTrimSeq.st ---- *)
(*
  Name: FB_DL_CoaterGapTrimSeq
  Category: DL_Process
  Version: 1.0.0
  Round: R90 / 2026-11-25
  开源溯源：clean-room 自研（族 锂电极片涂布辊压，ST 开源生态实测 0 命中，无外部代码引入）
  功能：1) 涂布间隙—面密度串级微调序：测厚稳定窗 → 算面密度相对偏差 → 点动间隙 → 稳定判定 →
           回到测厚（闭环迭代），偏差收敛到容差内即进换卷相并置完成位。
        2) 点动量算式采用「相对偏差 × 当前间隙」的比例律：面密度与湿膜厚度成正比，
           湿膜厚度与间隙成正比，故面密度相对偏差等于间隙相对偏差，
           修正量 Δgap = (实测 − 目标)/目标 × 当前间隙；该式量纲为 %/% × µm = µm，
           是无因次的相对量乘基准间隙，不需要额外的增益系数（增益已归一在比例律内部）。
        3) 每次点动量钳到 ±DL_JOG_MAX_UM，防止单次超大偏差把间隙一次拉穿；
           连续迭代次数受 DL_MAX_ITER 预算约束，超预算判「不收敛」故障而不是无限重试。
  边界条件：1) 非有限值闸：面密度实测、目标、间隙三路实值入参统一过
           NOT(x > -DL_BIG AND x < DL_BIG)，同时拦 NaN 与 Inf；命中即判信号无效（_bMeasOk=FALSE），
           在测厚相升级为「测厚信号丢失」故障，绝不把 NaN 送进偏差除法（R19）。
        2) 分母零闸：ABS(fArealTarget) > DL_EPS 才允许算相对偏差（目标为 0 时相对偏差无定义），
           目标为 0 或非有限在待机相直接判组态非法，禁止进入测量相。
        3) 时间零闸：tSettleS <= T#0S 时稳定窗定时器立即置 Q（等价于不做稳定判定）；
           这是合法组态（调试用），语义在此声明；同时另设 tonSettleOv 监视窗兜底。
        4) 间隙工艺闸：fGapUm 必须为正（间隙为 0 表示辊面接触，属设备危险状态），
           非正判组态非法并禁止启动。
        5) 相超时说明：eCgtMeasure 由 tonMeas 定时（测厚稳定窗）+ 非有限闸双重把关；
           eCgtJog 由 tonJog 定时；eCgtSettle 由 tonSettle 定时，并有 tonSettleOv 越限兜底；
           eCgtRollChange 为稳态持留相（等操作员撤令换卷），不设超时，设了会周期性误报；
           eCgtIdle / eCgtFault 为稳态相，同样不设超时。整序另设 tonSeq 总超时兜底。
        6) 状态机兜底：CASE 全态覆盖 + ELSE 强制回故障相；故障解除路径为
           (NOT xStart) AND (NOT xFault) AND 组态恢复，可达。
        7) FB 主体不使用 RETURN，统一单出口（跨平台可移植性）。
  量纲自证：fDevPct = (mg/cm2 − mg/cm2) / (mg/cm2) × 100 = 无因次 [%]；
           _fJogUm = ([%] / 100) × µm = µm，相对量乘基准间隙，量纲闭合；
           fGapCmdUm = µm + µm = µm，指令与实测间隙同量纲；tonXxx 的 PT 均为 [TIME]。
  码表 Error codes（本件格 0090_05xx，故障级一律 3 行内置 _uFault/_bFault/_eState）:
    16#0090_0501 故障级：组态非法（目标面密度/间隙/稳定时间越界或非有限）
    16#0090_0502 故障级：测厚信号丢失（面密度实测非有限）
    16#0090_0503 故障级：间隙微调不收敛（迭代次数超预算）
    16#0090_0504 故障级：稳定判定相超时（tonSettleOv 兜底命中）
    16#0090_0505 故障级：整序总超时
    16#0090_0506 故障级：外部故障输入 xFault
    16#0090_0507 故障级：状态机落 ELSE 兜底（非法相位 ID）
    16#0090_0508 信息级：单次点动量已饱和（达到 DL_JOG_MAX_UM，非故障）

  修订历史 Revision :
    2026-11-25  v1.0.0  R90 首版
*)

TYPE E_DL_CgtState :
(
    eCgtIdle       := 0,    // 待机：等启动上升沿 / Idle, awaiting start edge
    eCgtMeasure    := 10,   // 测厚：等稳定窗 / Measuring, awaiting stability window
    eCgtCalcDev    := 20,   // 算偏差：判收敛与迭代预算 / Deviation evaluation
    eCgtJog        := 30,   // 点动间隙：施加修正量 / Gap jog, applying correction
    eCgtSettle     := 40,   // 稳定判定：等涂层稳定 / Settling, awaiting stabilisation
    eCgtRollChange := 50,   // 换卷：完成保持，等撤令 / Roll change, done held until release
    eCgtFault      := 90    // 故障：锁存待解除 / Fault, latched awaiting release
);
END_TYPE

FUNCTION_BLOCK FB_DL_CoaterGapTrimSeq
VAR_INPUT
    xStart        : BOOL;    // 微调启动指令（上升沿有效）[bool] / Trim start command, edge triggered [bool]
    xFault        : BOOL;    // 外部故障汇总 [bool] / External fault aggregate [bool]
    fArealMeas    : REAL;    // 面密度实测值 [mg/cm2] / Measured areal loading [mg/cm2]
    fArealTarget  : REAL;    // 面密度目标值 [mg/cm2] / Target areal loading [mg/cm2]
    fGapUm        : REAL;    // 当前涂布间隙实测 [µm] / Current coating gap measurement [µm]
    tSettleS      : TIME;    // 稳定判定时长 [TIME] / Settling duration [TIME]
END_VAR
VAR_OUTPUT
    fGapCmdUm     : REAL;    // 间隙指令 [µm] / Gap command [µm]
    fDevPct       : REAL;    // 面密度相对偏差 [%] / Areal loading relative deviation [%]
    iIter         : INT;     // 已完成点动迭代次数 [-] / Completed jog iterations [-]
    xTrim         : BOOL;    // 正在微调（点动相）[bool] / Trimming active flag [bool]
    xDone         : BOOL;    // 微调完成保持位 [bool] / Trim complete held flag [bool]
    eState        : E_DL_CgtState;   // 状态出口，段尾单点映射 / State outlet, single-point mapped
    nErrId        : UDINT;   // 事件码，0 = 无事件 / Event code, 0 = none
END_VAR
VAR
    tonMeas       : TON;     // 测厚稳定窗定时 [TIME] / Measurement stability timer
    tonJog        : TON;     // 点动执行定时 [TIME] / Jog execution timer
    tonSettle     : TON;     // 稳定判定定时 [TIME] / Settling timer
    tonSettleOv   : TON;     // 稳定相越限兜底定时 [TIME] / Settling overrun watchdog timer
    tonSeq        : TON;     // 整序总超时定时 [TIME] / Whole-sequence timeout timer
    rtStart       : R_TRIG;  // 启动上升沿检测 [bool] / Start rising edge detector
    _eState       : E_DL_CgtState := E_DL_CgtState.eCgtIdle;   // 内部相位（CASE 唯一写入目标）
    _eStatePrev   : E_DL_CgtState := E_DL_CgtState.eCgtIdle;   // 上一拍相位快照（周期末更新）
    _bMeasOk      : BOOL;    // 测量链路有效性聚合 [bool] / Measurement chain validity aggregate
    _bCfgBad      : BOOL;    // 组态非法聚合 [bool] / Configuration invalid aggregate
    _bActive      : BOOL;    // 序激活（中间四相）[bool] / Sequence active flag [bool]
    _fDevRawPct   : REAL;    // 未饱和的相对偏差 [%] / Raw relative deviation [%]
    _fJogRawUm    : REAL;    // 未饱和的点动量 [µm] / Raw jog amount [µm]
    _fJogClampUm  : REAL;    // 饱和钳制后的点动量 [µm] / Clamped jog amount [µm]
    _fGapCmdLat   : REAL := 200.0;    // 间隙指令锁存（跨相保持；上电初值取安全张开位 200 µm，防冷启动输出 0 触发辊面接触）[µm]
    _iIter        : INT;     // 迭代次数内部量 [-] / Iteration counter internal [-]
    _bFault       : BOOL;    // 故障锁存位 [bool] / Latched fault flag [bool]
    _uInfo        : UDINT;   // 信息码，每拍重算 / Info code, recomputed every cycle
    _uFault       : UDINT;   // 故障码锁存 / Latched fault code
END_VAR
VAR CONSTANT
    DL_EPS        : REAL := 1.0E-9;      // 组态零闸阈值 [-] / Configuration zero gate threshold [-]
    DL_BIG        : REAL := 1.0E12;      // 非有限值闸量级上限 [-] / Finiteness gate magnitude [-]
    DL_PCT        : REAL := 100.0;       // 百分比换算因子 [%] / Percent conversion factor [%]
    DL_TOL_PCT    : REAL := 1.0;         // 面密度合格容差 [%] / Areal loading tolerance [%]
    DL_JOG_MAX_UM : REAL := 20.0;        // 单次点动饱和上限 [µm] / Single jog saturation limit [µm]
    DL_MAX_ITER   : INT  := 10;          // 迭代次数预算 [-] / Iteration budget [-]
    DL_MEASURE_S  : TIME := T#2S;        // 测厚稳定窗 [TIME] / Measurement stability window [TIME]
    DL_JOG_S      : TIME := T#1S;        // 点动执行时长 [TIME] / Jog execution duration [TIME]
    DL_OVER_MARGIN: TIME := T#10S;       // 稳定相越限兜底裕量 [TIME] / Settling watchdog margin [TIME]
    DL_SEQ_MAX    : TIME := T#10M;       // 整序总超时上限 [TIME] / Whole-sequence timeout [TIME]
END_VAR

(* —— 段 0：单拍量预清零（锁存量 _uFault/_bFault/_iIter/_fGapCmdLat/_eStatePrev 不入清单，R187①） —— *)
_uInfo := 16#0000_0000;                     // 信息码每拍重算 / Info code recomputed
nErrId := 16#0000_0000;                     // 事件码缺省无事件 / Event code defaults to none

(* —— 段 1：非有限值闸（R19：三路实值入参全覆盖，NaN 不得进入偏差除法） —— *)
_bMeasOk := (fArealMeas > -DL_BIG AND fArealMeas < DL_BIG)
            AND (fArealTarget > -DL_BIG AND fArealTarget < DL_BIG)
            AND (fGapUm > -DL_BIG AND fGapUm < DL_BIG);

(* —— 段 2：组态零闸（R4：目标面密度是偏差分母；间隙必须为正；稳定时长必须为正） —— *)
_bCfgBad := (NOT _bMeasOk)
            OR (ABS(fArealTarget) <= DL_EPS)                // 目标面密度不得为零
            OR (fGapUm <= DL_EPS)                           // 间隙必须为正（零间隙 = 辊面接触）
            OR (tSettleS <= T#0S);                          // 稳定时长必须为正（TIME 无法为 NaN）

(* —— 段 3：偏差与点动量解算（每拍重算，供观测与点动相直接取用） —— *)
IF _bCfgBad THEN
    _fDevRawPct := 0.0;                                 // 组态坏则偏差不计算，置 0
    _fJogRawUm := 0.0;                                  // 点动量置 0
ELSE
    _fDevRawPct := (fArealMeas - fArealTarget) / fArealTarget * DL_PCT;   // 实测 − 目标 [%]
    _fJogRawUm := (_fDevRawPct / DL_PCT) * fGapUm;      // 相对偏差 × 间隙 = 修正量 [µm]
END_IF
_fJogClampUm := LIMIT(-DL_JOG_MAX_UM, _fJogRawUm, DL_JOG_MAX_UM);          // 单次点动钳制 [µm]
IF ABS(_fJogRawUm) > DL_JOG_MAX_UM THEN
    _uInfo := 16#0090_0508;                             // 信息级：点动量已饱和（非故障）
END_IF

(* —— 段 4：激活量与定时器无条件周期刷新（R7：调用语句不得置于 IF/CASE 内） —— *)
_bActive := (_eState = E_DL_CgtState.eCgtMeasure) OR (_eState = E_DL_CgtState.eCgtCalcDev)
            OR (_eState = E_DL_CgtState.eCgtJog) OR (_eState = E_DL_CgtState.eCgtSettle);
rtStart(CLK := xStart);                                                     // 启动上升沿，每拍必调
tonMeas(IN := (_eState = E_DL_CgtState.eCgtMeasure), PT := DL_MEASURE_S);   // 测厚稳定窗
tonJog(IN := (_eState = E_DL_CgtState.eCgtJog), PT := DL_JOG_S);            // 点动执行时长
tonSettle(IN := (_eState = E_DL_CgtState.eCgtSettle), PT := tSettleS);      // 稳定判定定时
tonSettleOv(IN := (_eState = E_DL_CgtState.eCgtSettle),
            PT := tSettleS + DL_OVER_MARGIN);                               // 稳定相越限兜底
tonSeq(IN := _bActive, PT := DL_SEQ_MAX);                                    // 整序总超时

(* —— 段 5：全局故障拦截（优先级最高；已锁存则不再改写码值，禁同拍抹除） —— *)
IF xFault AND (NOT _bFault) THEN
    _uFault := 16#0090_0506;                // 故障级：外部故障输入
    _bFault := TRUE;                        // 锁存（3 行内置，R45 配对）
    _eState := E_DL_CgtState.eCgtFault;
END_IF
IF (NOT _bMeasOk) AND (_bActive) AND (NOT _bFault) THEN
    _uFault := 16#0090_0502;                // 故障级：测厚信号丢失
    _bFault := TRUE;                        // 锁存
    _eState := E_DL_CgtState.eCgtFault;
END_IF
IF tonSeq.Q AND _bActive AND (NOT _bFault) THEN
    _uFault := 16#0090_0505;                // 故障级：整序总超时
    _bFault := TRUE;                        // 锁存
    _eState := E_DL_CgtState.eCgtFault;
END_IF
IF _bCfgBad AND (NOT _bFault) AND (_eState <> E_DL_CgtState.eCgtIdle) THEN
    _uFault := 16#0090_0501;                // 故障级：组态非法
    _bFault := TRUE;                        // 锁存
    _eState := E_DL_CgtState.eCgtFault;
END_IF

(* —— 段 6：相位机（只做迁移；出口在段 8 单点映射） —— *)
CASE _eState OF

E_DL_CgtState.eCgtIdle:
    IF NOT xStart THEN
        ;                                   // 等启动，撤令状态保持 / Waiting for start
    ELSIF _bCfgBad THEN
        _uFault := 16#0090_0501;            // 故障级：组态非法（启动前置校验）
        _bFault := TRUE;
        _eState := E_DL_CgtState.eCgtFault;
    ELSIF rtStart.Q THEN
        _eState := E_DL_CgtState.eCgtMeasure;   // 新序开始：进测厚相（迭代预算在段 7 清零）
    END_IF

E_DL_CgtState.eCgtMeasure:
    IF NOT xStart THEN
        _eState := E_DL_CgtState.eCgtIdle;      // 撤令：回待机
    ELSIF tonMeas.Q THEN
        _eState := E_DL_CgtState.eCgtCalcDev;   // 稳定窗结束：进算偏差相
    END_IF

E_DL_CgtState.eCgtCalcDev:
    IF NOT xStart THEN
        _eState := E_DL_CgtState.eCgtIdle;
    ELSIF ABS(_fDevRawPct) <= DL_TOL_PCT THEN
        _eState := E_DL_CgtState.eCgtRollChange;    // 本拍合法事件（已收敛）优先（R275）
    ELSIF _iIter >= DL_MAX_ITER THEN
        _uFault := 16#0090_0503;            // 故障级：迭代超预算，不收敛
        _bFault := TRUE;
        _eState := E_DL_CgtState.eCgtFault;
    ELSE
        _eState := E_DL_CgtState.eCgtJog;   // 未收敛且预算内：进点动相
    END_IF

E_DL_CgtState.eCgtJog:
    IF NOT xStart THEN
        _eState := E_DL_CgtState.eCgtIdle;
    ELSIF tonJog.Q THEN
        _eState := E_DL_CgtState.eCgtSettle;    // 点动完成：进稳定判定相
    END_IF

E_DL_CgtState.eCgtSettle:
    IF NOT xStart THEN
        _eState := E_DL_CgtState.eCgtIdle;
    ELSIF tonSettle.Q THEN
        _eState := E_DL_CgtState.eCgtMeasure;   // 稳定：回测厚，闭环复测
    ELSIF tonSettleOv.Q THEN
        _uFault := 16#0090_0504;            // 故障级：稳定相越限兜底命中
        _bFault := TRUE;
        _eState := E_DL_CgtState.eCgtFault;
    END_IF

E_DL_CgtState.eCgtRollChange:
    IF xFault THEN
        _uFault := 16#0090_0506;            // 故障级：换卷相外部故障
        _bFault := TRUE;
        _eState := E_DL_CgtState.eCgtFault;
    ELSIF NOT xStart THEN
        _eState := E_DL_CgtState.eCgtIdle;  // 撤令：回待机，完成位在段 7 清
    END_IF

E_DL_CgtState.eCgtFault:
    IF (NOT xStart) AND (NOT xFault) AND (NOT _bCfgBad) THEN
        _bFault := FALSE;                   // 解除路径：撤令 + 外部故障消失 + 组态恢复（可达）
        _uFault := 16#0000_0000;            // 清锁存码
        _eState := E_DL_CgtState.eCgtIdle;  // 回待机
    END_IF

ELSE
    _uFault := 16#0090_0507;                // 故障级：非法相位 ID 兜底
    _bFault := TRUE;                        // 锁存
    _eState := E_DL_CgtState.eCgtFault;     // 强制回故障相

END_CASE

(* —— 段 7：后置段（R23：迭代预算、间隙指令锁存、快照统一放在迁移判断之后） —— *)
IF (_eState = E_DL_CgtState.eCgtMeasure) AND (_eStatePrev = E_DL_CgtState.eCgtIdle) THEN
    _iIter := 0;                            // 新序开始：迭代预算清零（禁跨相重试预算不清零）
END_IF
IF (_eState = E_DL_CgtState.eCgtJog) AND (_eStatePrev = E_DL_CgtState.eCgtCalcDev) THEN
    _iIter := _iIter + 1;                   // 进入点动即消耗一次迭代预算
END_IF

IF _eState = E_DL_CgtState.eCgtJog THEN
    _fGapCmdLat := LIMIT(DL_EPS, fGapUm + _fJogClampUm, DL_BIG);   // 点动相：实测间隙 + 修正量
ELSIF (NOT _bActive) AND _bMeasOk AND (NOT _bCfgBad) THEN
    _fGapCmdLat := LIMIT(DL_EPS, fGapUm, DL_BIG);   // 非激活相：指令跟随实测（仅测量有效时）
ELSIF NOT _bActive THEN
    ;                                   // 测量无效/组态非法：保持上拍指令，不复制 NaN 实测值
END_IF

_eStatePrev := _eState;                     // 快照统一在周期末尾更新（R23）

(* —— 段 8：出口单点映射（名实同源；指令/标志由状态与锁存导出，不在多分支各写一遍） —— *)
fGapCmdUm := _fGapCmdLat;                                       // 间隙指令出口 [µm]
fDevPct := LIMIT(-DL_BIG, _fDevRawPct, DL_BIG);                 // 偏差出口（已闸非有限）
iIter := _iIter;                                                // 迭代次数出口
xTrim := (_eState = E_DL_CgtState.eCgtJog) AND (NOT _bFault);   // 微调中出口
xDone := (_eState = E_DL_CgtState.eCgtRollChange) AND (NOT _bFault);   // 完成位出口
eState := _eState;                                              // 状态出口单点映射
IF _bFault THEN
    nErrId := _uFault;                      // 故障锁存码回放（不在故障相按当下输入重推断）
ELSE
    nErrId := _uInfo;                       // 信息码
END_IF

END_FUNCTION_BLOCK

(* ---- FB_DL_CoatingGapMeasure.st ---- *)
// =====================================================================
// FB_DL_CoatingGapMeasure.st
// 涂布留白（Gap）宽度与边缘对齐判定（像素到毫米标定 + 区间带 + 窗口一致性）
// Coating gap width judge with pixel calibration and band check
// 所属子库: DL_Process    版本: v1.0.0    兼容: CODESYS V3.5+ / TwinCAT 3 / 汇川 InoProShop
// 码位: 16#0005_048A ~ 16#0005_048E (本件独占 5 槽, 勿复用)
// 溯源: 道莅 clean-room 防御性实现
//       来源组标签: lithium-battery, coating, vision-metrology, tolerance
// 修改记录: R30 初版 (ROUND_PLAN_R30 序 13)
// 分层声明: 带判定消费 DL_Base 的 FC_DL_IntervalMembership（双闭组合,
//           恰好落在带端点判带内）; 窗口一致性消费 DL_MathData 的
//           FB_DL_SignalStatistics（窗口均值/极差经引脚注入, 本件不重写统计）
// =====================================================================
FUNCTION_BLOCK FB_DL_CoatingGapMeasure
VAR_INPUT
    afPixEdge1    : REAL := 0.0;    // 第一边缘像素坐标 / First edge pixel coordinate [px]
    afPixEdge2    : REAL := 0.0;    // 第二边缘像素坐标 / Second edge pixel coordinate [px]
    fPixToMm      : REAL := 0.01;   // 标定系数 0~10 mm/px / Calibration factor [mm/px]
    afGapLo_mm    : REAL := 8.0;    // 留白带下限 0~100 mm / Gap band lower [mm]
    afGapHi_mm    : REAL := 12.0;   // 留白带上限 0~100 mm / Gap band upper [mm]
    fWinTolPct    : REAL := 10.0;   // 窗口一致性容差（相对带宽）0~100 百分比 / Window consistency tolerance [pct]
    uWinSize      : USINT := 8;     // 窗口样本数配置（传给上游统计件）2~256 / Window size config
    fWinMean_mm   : REAL := 0.0;    // 窗口均值注入（统计件 fMean 语义）/ Window mean injected [mm]
    fWinRange_mm  : REAL := 0.0;    // 窗口极差注入（统计件 fRange 语义）/ Window range injected [mm]
    bWinStatValid : BOOL := FALSE;  // 窗口统计有效注入（统计件 bValid 语义）/ Window stat valid injected
END_VAR
VAR_OUTPUT
    fGap_mm         : REAL  := 0.0;   // 留白宽度 / Gap width [mm]
    bGapOk          : BOOL  := FALSE; // 带内判定 / In-band flag
    bWindowConsist  : BOOL  := FALSE; // 窗口一致性 / Window consistency flag
    eErr            : UDINT := 16#0005_048A;  // 错误码 / Error code
END_VAR
VAR
    bCfgErr    : BOOL  := FALSE;      // 组态非法标记 / Configuration error flag
    bSnsErr    : BOOL  := FALSE;      // 传感器故障标记（边缘序颠倒）/ Sensor error flag
    fBandSpan  : REAL  := 0.0;        // 带宽 / Band span [mm]
    bInBand    : BOOL  := FALSE;      // 区间判定返回 / Interval membership return
    fGapL      : LREAL := 0.0;        // 留白宽度双精度临时量 / Gap width LREAL temporary [mm]
    fLoL       : LREAL := 0.0;        // 带下限双精度临时量 / Band lower LREAL temporary [mm]
    fHiL       : LREAL := 0.0;        // 带上限双精度临时量 / Band upper LREAL temporary [mm]
END_VAR

// ---------------------------------------------------------------------
// 代码位表（本件独占, 勿复用）:
//   16#0005_048A 信息 留白判定正常（带内且窗口一致性满足）
//   16#0005_048B 信息 留白越带（带外, 判定值仍逐拍输出）
//   16#0005_048C 故障 组态非法（标定系数非有限或不大于 0, 带倒置, 容差越域,
//                窗口样本数小于 2）; 解除式 = 恢复合法组态
//   16#0005_048D 故障 边缘序颠倒（第二边缘不大于第一边缘 → 负留白, 传感器故障）,
//                解除式 = 边缘序恢复正差
//   16#0005_048E 信息 窗口一致性不满足（均值/极差注入超容差或统计无效）
// ---------------------------------------------------------------------

// ---- 组态闸 / Configuration gate ----
bCfgErr := FALSE;                   // 组态标记复位 / Reset config flag
IF (fPixToMm <> fPixToMm) OR (fPixToMm <= 0.0) OR (fPixToMm > 10.0) THEN
    bCfgErr := TRUE;                // 标定系数非法 / Illegal calibration
END_IF
IF (afGapLo_mm <> afGapLo_mm) OR (afGapHi_mm <> afGapHi_mm)
   OR (afGapHi_mm < afGapLo_mm) THEN
    bCfgErr := TRUE;                // 带非法或倒置 / Illegal or inverted band
END_IF
IF (fWinTolPct <> fWinTolPct) OR (fWinTolPct < 0.0) OR (fWinTolPct > 100.0) THEN
    bCfgErr := TRUE;                // 容差越域 / Illegal tolerance
END_IF
IF uWinSize < 2 THEN
    bCfgErr := TRUE;                // 窗口过小, 统计无意义 / Window too small
END_IF

// ---- 输出缺省收口 / Output defaults ----
fGap_mm := 0.0;                     // 缺省零 / Default zero
bGapOk := FALSE;                    // 缺省带外 / Default out of band
bWindowConsist := FALSE;            // 缺省不一致 / Default inconsistent
bSnsErr := FALSE;                   // 传感器标记复位 / Reset sensor flag

IF NOT bCfgErr THEN
    IF (afPixEdge1 <> afPixEdge1) OR (ABS(afPixEdge1) >= 1.0E12)
       OR (afPixEdge2 <> afPixEdge2) OR (ABS(afPixEdge2) >= 1.0E12) THEN
        bSnsErr := TRUE;            // 边缘坐标非有限 / Non-finite edge coordinate
    ELSE
        fGap_mm := (afPixEdge2 - afPixEdge1) * fPixToMm;    // 像素差换算毫米 / Pixel diff to mm
        IF fGap_mm < 0.0 THEN
            bSnsErr := TRUE;        // 边缘序颠倒判负留白 / Reversed edges, negative gap
        ELSE
            // 带判定消费区间判定函数（双闭组合, 端点恰落判带内）/ Band via interval membership
            fGapL := REAL_TO_LREAL(fGap_mm);
            fLoL  := REAL_TO_LREAL(afGapLo_mm);
            fHiL  := REAL_TO_LREAL(afGapHi_mm);
            bInBand := FC_DL_IntervalMembership(fGapL, fLoL, fHiL,
                        E_DL_IntervalKind.eClosedClosed, 1.0E-9);
            bGapOk := bInBand;      // 带内判定 / In-band result
            // 窗口一致性消费注入统计量（不重写统计）/ Window consistency via injected stats
            fBandSpan := afGapHi_mm - afGapLo_mm;   // 带宽 / Band span [mm]
            IF bWinStatValid AND (fWinMean_mm = fWinMean_mm) AND (fWinRange_mm = fWinRange_mm) THEN
                bWindowConsist := (ABS(fWinMean_mm - fGap_mm) <= (fBandSpan * fWinTolPct / 100.0))
                               AND (fWinRange_mm <= (2.0 * fBandSpan * fWinTolPct / 100.0));
            ELSE
                bWindowConsist := FALSE;    // 统计无效或注入非有限判不一致 / Invalid stats judged inconsistent
            END_IF
        END_IF
    END_IF
END_IF

// ---- 错误码仲裁 / Error arbitration ----
IF bCfgErr THEN
    eErr := 16#0005_048C;           // 组态非法 / Config fault
ELSIF bSnsErr THEN
    eErr := 16#0005_048D;           // 边缘序颠倒 / Reversed edges
ELSIF NOT bGapOk THEN
    eErr := 16#0005_048B;           // 留白越带 / Out of band
ELSIF NOT bWindowConsist THEN
    eErr := 16#0005_048E;           // 窗口一致性不满足 / Window inconsistent
ELSE
    eErr := 16#0005_048A;           // 判定正常 / Judgement normal
END_IF

END_FUNCTION_BLOCK

(* ---- FB_DL_CoinCellAssembler.st ---- *)
(*
  ==================================================================
  组件名 Component  : FB_DL_CoinCellAssembler
  分类   Category   : DL_Process
  版本   Version    : 1.0.1
  功能   Purpose    : 扣电组装工站模板（叠片 — 压紧 — 封口）。以 ENUM + CASE 相位机
                      编排七相：空闲 → 上料 → 叠片 → 压紧 → 封口 → 下料 → 完成；
                      每相输出本相命令并等本相就绪信号，各相独立超时（独立成因码，
                      R190 归因唯一）；压紧相另设压力上限保护，超限立即跳故障相。
                      完成相出单拍周期完成脉冲并累加周期计数。
  溯源   Origin     : 扣电组装（叠片 / 压紧 / 封口）为通用小电芯工站时序语义；本件为
                      clean-room 实现，仅借鉴来源分类与参数域组织（来源标签
                      roadmap-p2-coincell），道莅原创设计，未复制任何闭源代码行。
  平台   Platform   : 纯 IEC 61131-3（TON / R_TRIG / REAL 运算，无私有库）
  作者   Author     : 道莅代码库 · PLC 编程专家（R55）
  ------------------------------------------------------------------
  同拍多窗说明（R100）：五个超时窗互斥 —— 每窗的 IN 均串「本相」闸，任一时刻只有一个
                      窗在计时，因此不存在同拍双窗配比约束；若后续改为并行工位，必须补
                      配比约束句后再改 IN 结构。
  边界 Boundary     :
                      一 本件只出工站级相命令与就绪判据，不驱动伺服 / 气缸本体（属主边界）；
                      二 每相命令只在对应相位为真，相外一律撤除（每拍预置撤除）；
                      三 五个超时件全部无条件周期刷新，IN 串相位闸与故障闸（禁分支内调用）；
                      四 压力上限保护独立成码，不与超时码合并（R190）；
                      五 无全局变量、无外部变量声明、无物理地址寻址。
  输出契约 Output contract:
                      五个命令出口为「相位派生电平」，相外恒假；
                      bCycleDone 为单拍脉冲（内部位置置位、统一出口映射后撤销）；
                      nCycleCnt 只在下料就绪那一拍递增，饱和到上限；
                      eCause 故障级成因与 bError 配对（R45），信息级永不置 bError。
  修订记录 Revision  :
    2026-11-20  v1.0.0  R55 首版（批 4 · 序号 18）
    2026-11-20  v1.0.1  R56 返修（7.3）：删除死变量 _eCause（信息级成因全文件无任何
                        写入路径、恒为 eNone），段 7 出口简化为故障级成因锁存直映。
  ==================================================================
*)

TYPE E_DL_CcaPhase :
(
    eIdle   := 0,       // 空闲：等启动沿 / idle, waiting for the start edge
    eLoad   := 10,      // 上料：等上料就绪 / loading, waiting for the load ready signal
    eStack  := 20,      // 叠片：等叠片就绪 / stacking, waiting for the stack ready signal
    ePress  := 30,      // 压紧：等压紧就绪（含压力上限保护）/ pressing, waiting for the press ready signal with force protection
    eSeal   := 40,      // 封口：等封口就绪 / sealing, waiting for the seal ready signal
    eUnload := 50,      // 下料：等下料就绪 / unloading, waiting for the unload ready signal
    eDone   := 60,      // 完成：周期完成脉冲已出，驻留一拍以上 / done, the cycle pulse has been raised
    eFault  := 90       // 故障：成因锁存 / fault, the cause is latched
);
END_TYPE

TYPE E_DL_CcaCause :
(
    eNone       := 0,   // 无成因 / no cause
    eCfgIllegal := 1,   // 组态非法：时间或力量程越域（故障级，与 bError 配对）/ illegal config, time or force range out of domain
    eLoadTo     := 2,   // 上料超时（故障级，与 bError 配对）/ load timeout, a fault paired with bError
    eStackTo    := 3,   // 叠片超时（故障级，与 bError 配对）/ stack timeout, a fault paired with bError
    ePressTo    := 4,   // 压紧超时（故障级，与 bError 配对）/ press timeout, a fault paired with bError
    eSealTo     := 5,   // 封口超时（故障级，与 bError 配对）/ seal timeout, a fault paired with bError
    eUnloadTo   := 6,   // 下料超时（故障级，与 bError 配对）/ unload timeout, a fault paired with bError
    eForceOver  := 7    // 压紧力越上限（故障级，与 bError 配对）/ press force above the ceiling, a fault paired with bError
);
END_TYPE

FUNCTION_BLOCK FB_DL_CoinCellAssembler
VAR_INPUT
    bEnable      : BOOL := TRUE;             // 使能，失能时撤命令回空闲 [-] / enable, disabling withdraws the commands and returns to idle
    bReset       : BOOL := FALSE;           // 复位上升沿清故障锁存并回空闲 [-] / reset rising edge clears the fault latch and returns to idle
    bStart       : BOOL := FALSE;            // 周期启动脉冲，上升沿受理 [-] / cycle start pulse, accepted on the rising edge
    bLoadOk      : BOOL := FALSE;            // 上料就绪（物料到位）[-] / load ready, the part is in place
    bStackOk     : BOOL := FALSE;            // 叠片就绪（叠片数达标）[-] / stack ready, the layer count is reached
    bPressOk     : BOOL := FALSE;            // 压紧就绪（压力到位）[-] / press ready, the force is reached
    bSealOk      : BOOL := FALSE;            // 封口就绪（封口完成信号）[-] / seal ready
    bUnloadOk    : BOOL := FALSE;            // 下料就绪（物料已取出）[-] / unload ready, the part was removed
    fPressForceN : REAL := 0.0;              // 压紧力实测 [牛顿] / measured press force [newton]
    fPressMaxN   : REAL := 5000.0;           // 压紧力上限 [牛顿]，域 大于零 / press force ceiling [newton], domain above zero
    tLoadTo      : TIME := T#15S;            // 上料超时 [毫秒]，域 大于零 / load timeout [millisecond], domain above zero
    tStackTo     : TIME := T#60S;            // 叠片超时 [毫秒]，域 大于零 / stack timeout [millisecond], domain above zero
    tPressTo     : TIME := T#30S;            // 压紧超时 [毫秒]，域 大于零 / press timeout [millisecond], domain above zero
    tSealTo      : TIME := T#30S;            // 封口超时 [毫秒]，域 大于零 / seal timeout [millisecond], domain above zero
    tUnloadTo    : TIME := T#15S;            // 下料超时 [毫秒]，域 大于零 / unload timeout [millisecond], domain above zero
END_VAR
VAR_OUTPUT
    bLoadCmd     : BOOL := FALSE;            // 上料相命令 [-] / load phase command
    bStackCmd    : BOOL := FALSE;            // 叠片相命令 [-] / stack phase command
    bPressCmd    : BOOL := FALSE;            // 压紧相命令 [-] / press phase command
    bSealCmd     : BOOL := FALSE;            // 封口相命令 [-] / seal phase command
    bUnloadCmd   : BOOL := FALSE;            // 下料相命令 [-] / unload phase command
    bCycleDone   : BOOL := FALSE;            // 周期完成单拍脉冲 [-] / cycle done single-shot pulse
    bBusy        : BOOL := FALSE;            // 工站忙（非空闲非故障）[-] / station busy, neither idle nor faulted
    nCycleCnt    : UDINT := 0;               // 周期完成计数（饱和到上限）[次] / completed cycle count, saturated [cycle]
    ePhase       : E_DL_CcaPhase := E_DL_CcaPhase.eIdle; // 相位出口 [枚举] / phase outlet [enum]
    eCause       : E_DL_CcaCause := E_DL_CcaCause.eNone; // 成因出口 [枚举] / cause outlet [enum]
    bError       : BOOL := FALSE;            // 故障锁存标志 [-] / fault latch flag
END_VAR
VAR
    rtStart      : R_TRIG;                   // 启动沿检测，段 0 无条件刷新 / start edge detector, refreshed unconditionally in segment zero
    rtReset      : R_TRIG;                   // 复位沿检测，段 0 无条件刷新 / reset edge detector, refreshed unconditionally in segment zero
    tonLoad      : TON;                      // 上料超时，段 0 无条件刷新 / load timeout, refreshed unconditionally in segment zero
    tonStack     : TON;                      // 叠片超时，段 0 无条件刷新 / stack timeout, refreshed unconditionally in segment zero
    tonPress     : TON;                      // 压紧超时，段 0 无条件刷新 / press timeout, refreshed unconditionally in segment zero
    tonSeal      : TON;                      // 封口超时，段 0 无条件刷新 / seal timeout, refreshed unconditionally in segment zero
    tonUnload    : TON;                      // 下料超时，段 0 无条件刷新 / unload timeout, refreshed unconditionally in segment zero
    _ePhase      : E_DL_CcaPhase := E_DL_CcaPhase.eIdle;  // 内部相位，CASE 唯一写入目标 / internal phase, the only CASE write target
    _eFaultCause : E_DL_CcaCause := E_DL_CcaCause.eNone;  // 故障级成因，锁存至复位沿（本件全部成因均为故障级，信息级死变量 _eCause 已于 R56 删除）/ fault cause, latched until the reset edge, every cause here is fault grade
    _bFault      : BOOL := FALSE;            // 故障锁存位 [-] / fault latch bit
    _bInit       : BOOL := FALSE;            // 首扫初始化完成标志（R310）/ first scan initialisation flag
    _bCfgBad     : BOOL := FALSE;            // 组态非法判定 [-] / illegal configuration verdict
    _bDoneInt    : BOOL := FALSE;            // 周期完成脉冲内部位，统一出口映射 / internal cycle done bit, mapped at the unified outlet
    _bForceOk    : BOOL := FALSE;            // 压紧力域闸通过 [-] / press force domain gate passed
    _nCycle      : UDINT := 0;               // 周期计数工作值 [次] / cycle count working value [cycle]
END_VAR
VAR CONSTANT
    DL_CCA_FORCE_MAX : REAL := 1.0E7;        // 压紧力量级上限 [牛顿] / press force magnitude ceiling [newton]
    DL_CCA_CYCLE_MAX : UDINT := 2000000000;  // 周期计数饱和上限（常量在 DINT 可表范围内）[次] / cycle count saturation ceiling, the constant fits in DINT
END_VAR

// 段 0｜定时器与沿检测无条件周期刷新（禁入分支），IN 只串相位闸与故障闸（R212）/ segment 0, unconditional refresh with phase and fault gates on IN only
rtStart(CLK := bStart); // 启动沿无条件刷新 / unconditional refresh of the start edge
rtReset(CLK := bReset); // 复位沿无条件刷新 / unconditional refresh of the reset edge
tonLoad(IN := (_ePhase = E_DL_CcaPhase.eLoad) AND (NOT _bFault), PT := tLoadTo); // 上料超时 / load timeout
tonStack(IN := (_ePhase = E_DL_CcaPhase.eStack) AND (NOT _bFault), PT := tStackTo); // 叠片超时 / stack timeout
tonPress(IN := (_ePhase = E_DL_CcaPhase.ePress) AND (NOT _bFault), PT := tPressTo); // 压紧超时 / press timeout
tonSeal(IN := (_ePhase = E_DL_CcaPhase.eSeal) AND (NOT _bFault), PT := tSealTo); // 封口超时 / seal timeout
tonUnload(IN := (_ePhase = E_DL_CcaPhase.eUnload) AND (NOT _bFault), PT := tUnloadTo); // 下料超时 / unload timeout

// 段 1｜首扫初始化（R310）/ segment 1, first scan initialisation
IF NOT _bInit THEN // 首扫一拍 / the very first scan
    _bInit := TRUE; // 置首扫完成标志 / raise the first scan flag
    _ePhase := E_DL_CcaPhase.eIdle; // 相位从空闲起步 / the phase starts from idle
    _eFaultCause := E_DL_CcaCause.eNone; // 故障级成因清零 / clear the fault cause
    _bFault := FALSE; // 故障锁存清零 / clear the fault latch
    _nCycle := 0; // 周期计数清零 / clear the cycle count
END_IF

// 段 2｜复位沿作用域：清锁存 / 迁相位 / 清脉冲内部位（计数不清，属产量资产）/ segment 2, reset edge scope
IF rtReset.Q THEN // 复位沿 / reset edge
    _bFault := FALSE; // 作用域一：清故障锁存 / scope one, clear the fault latch
    _eFaultCause := E_DL_CcaCause.eNone; // 作用域一：清故障级成因 / scope one, clear the fault cause
    _ePhase := E_DL_CcaPhase.eIdle; // 作用域二：迁回空闲相 / scope two, migrate back to idle
    _bDoneInt := FALSE; // 作用域二：清周期完成脉冲内部位 / scope two, clear the internal cycle done bit
END_IF

// 段 3｜组态域闸（R151 全覆盖）：五个时间引脚与力量程 / segment 3, configuration domain gate over every pin
_bCfgBad := FALSE; // 组态非法预置假 / preset the illegal configuration verdict to false
IF (tLoadTo <= T#0S) OR (tStackTo <= T#0S) OR (tPressTo <= T#0S) OR (tSealTo <= T#0S) OR (tUnloadTo <= T#0S) THEN // 时间引脚非正 / a time pin is not positive
    _bCfgBad := TRUE; // 判非法 / mark illegal
END_IF
IF (fPressMaxN <= 0.0) OR (fPressMaxN <> fPressMaxN) OR (fPressMaxN > DL_CCA_FORCE_MAX) THEN // 力量程越域 / the force range is out of domain
    _bCfgBad := TRUE; // 判非法 / mark illegal
END_IF
IF _bCfgBad AND (NOT _bFault) THEN // 组态非法且未锁存 / illegal configuration and not yet latched
    _bFault := TRUE; // 置故障锁存 / raise the fault latch
    _eFaultCause := E_DL_CcaCause.eCfgIllegal; // 故障级成因 (R45 配对 bError) / fault grade cause paired with bError
    _ePhase := E_DL_CcaPhase.eFault; // 迁故障相 / migrate to the fault phase
END_IF

// 段 4｜命令预置与压紧力闸：命令为相位派生电平，每拍先撤除 / segment 4, command preset and press force gate
bLoadCmd := FALSE; // 上料命令预置撤除 / preset the load command withdrawn
bStackCmd := FALSE; // 叠片命令预置撤除 / preset the stack command withdrawn
bPressCmd := FALSE; // 压紧命令预置撤除 / preset the press command withdrawn
bSealCmd := FALSE; // 封口命令预置撤除 / preset the seal command withdrawn
bUnloadCmd := FALSE; // 下料命令预置撤除 / preset the unload command withdrawn
_bForceOk := (fPressForceN = fPressForceN) AND ((fPressForceN - fPressForceN) = (fPressForceN - fPressForceN)) AND (fPressForceN <= fPressMaxN); // 压紧力有限且不越上限 / the press force is finite and within the ceiling

// 段 5｜相位机：ENUM + CASE，含 ELSE 非法相位兜底（R128）/ segment 5, phase machine with an ELSE fallback for illegal phases
CASE _ePhase OF
E_DL_CcaPhase.eIdle: // 空闲相：等启动沿 / idle, waiting for the start edge
    IF rtStart.Q AND bEnable AND (NOT _bFault) THEN // 启动沿且使能无故障 / start edge while enabled and unfaulted
        _ePhase := E_DL_CcaPhase.eLoad; // 迁上料相 / migrate to the load phase
    END_IF

E_DL_CcaPhase.eLoad: // 上料相：命令自锁于本相 / load phase, the command lives inside this phase
    bLoadCmd := TRUE; // 出上料命令 / raise the load command
    IF bLoadOk THEN // 上料就绪 / load ready
        _ePhase := E_DL_CcaPhase.eStack; // 迁叠片相 / migrate to the stack phase
    ELSIF tonLoad.Q THEN // 上料超时 / load timed out
        _bFault := TRUE; // 置故障锁存 / raise the fault latch
        _eFaultCause := E_DL_CcaCause.eLoadTo; // 故障级成因（独立码，R45 配对 bError）/ independent fault code paired with bError
        _ePhase := E_DL_CcaPhase.eFault; // 迁故障相 / migrate to the fault phase
    END_IF

E_DL_CcaPhase.eStack: // 叠片相 / stack phase
    bStackCmd := TRUE; // 出叠片命令 / raise the stack command
    IF bStackOk THEN // 叠片就绪 / stack ready
        _ePhase := E_DL_CcaPhase.ePress; // 迁压紧相 / migrate to the press phase
    ELSIF tonStack.Q THEN // 叠片超时 / stack timed out
        _bFault := TRUE; // 置故障锁存 / raise the fault latch
        _eFaultCause := E_DL_CcaCause.eStackTo; // 故障级成因（独立码）/ independent fault code
        _ePhase := E_DL_CcaPhase.eFault; // 迁故障相 / migrate to the fault phase
    END_IF

E_DL_CcaPhase.ePress: // 压紧相：命令 + 压力上限保护双判 / press phase with force protection
    bPressCmd := TRUE; // 出压紧命令 / raise the press command
    IF NOT _bForceOk THEN // 压紧力越上限或非有限 / the force is above the ceiling or non-finite
        _bFault := TRUE; // 置故障锁存 / raise the fault latch
        _eFaultCause := E_DL_CcaCause.eForceOver; // 故障级成因（独立码，不与超时合并）/ independent fault code, never merged with a timeout
        _ePhase := E_DL_CcaPhase.eFault; // 迁故障相 / migrate to the fault phase
    ELSIF bPressOk THEN // 压紧就绪 / press ready
        _ePhase := E_DL_CcaPhase.eSeal; // 迁封口相 / migrate to the seal phase
    ELSIF tonPress.Q THEN // 压紧超时 / press timed out
        _bFault := TRUE; // 置故障锁存 / raise the fault latch
        _eFaultCause := E_DL_CcaCause.ePressTo; // 故障级成因（独立码）/ independent fault code
        _ePhase := E_DL_CcaPhase.eFault; // 迁故障相 / migrate to the fault phase
    END_IF

E_DL_CcaPhase.eSeal: // 封口相 / seal phase
    bSealCmd := TRUE; // 出封口命令 / raise the seal command
    IF bSealOk THEN // 封口就绪 / seal ready
        _ePhase := E_DL_CcaPhase.eUnload; // 迁下料相 / migrate to the unload phase
    ELSIF tonSeal.Q THEN // 封口超时 / seal timed out
        _bFault := TRUE; // 置故障锁存 / raise the fault latch
        _eFaultCause := E_DL_CcaCause.eSealTo; // 故障级成因（独立码）/ independent fault code
        _ePhase := E_DL_CcaPhase.eFault; // 迁故障相 / migrate to the fault phase
    END_IF

E_DL_CcaPhase.eUnload: // 下料相 / unload phase
    bUnloadCmd := TRUE; // 出下料命令 / raise the unload command
    IF bUnloadOk THEN // 下料就绪 / unload ready
        IF _nCycle < DL_CCA_CYCLE_MAX THEN // 计数未达饱和上限 / below the saturation ceiling
            _nCycle := _nCycle + 1; // 周期计数递增 / increment the cycle count
        END_IF
        _bDoneInt := TRUE; // 周期完成脉冲内部位置位（统一出口映射，R187）/ raise the internal cycle done bit, mapped at the unified outlet
        _ePhase := E_DL_CcaPhase.eDone; // 迁完成相 / migrate to the done phase
    ELSIF tonUnload.Q THEN // 下料超时 / unload timed out
        _bFault := TRUE; // 置故障锁存 / raise the fault latch
        _eFaultCause := E_DL_CcaCause.eUnloadTo; // 故障级成因（独立码）/ independent fault code
        _ePhase := E_DL_CcaPhase.eFault; // 迁故障相 / migrate to the fault phase
    END_IF

E_DL_CcaPhase.eDone: // 完成相：驻留，等复位或新启动 / done phase, held until reset or a new start
    IF rtStart.Q AND bEnable THEN // 新启动沿 / a new start edge
        _ePhase := E_DL_CcaPhase.eLoad; // 重启上料相 / restart from the load phase
    END_IF

E_DL_CcaPhase.eFault: // 故障相：全撤命令，等复位沿 / fault phase with all commands withdrawn
    bLoadCmd := FALSE; // 撤上料命令 / withdraw the load command
    bStackCmd := FALSE; // 撤叠片命令 / withdraw the stack command
    bPressCmd := FALSE; // 撤压紧命令 / withdraw the press command
    bSealCmd := FALSE; // 撤封口命令 / withdraw the seal command
    bUnloadCmd := FALSE; // 撤下料命令 / withdraw the unload command

ELSE // 非法相位兜底（R128）/ illegal phase fallback
    _bFault := TRUE; // 置故障锁存 / raise the fault latch
    _eFaultCause := E_DL_CcaCause.eCfgIllegal; // 故障级成因记组态非法 / record the illegal configuration cause
    _ePhase := E_DL_CcaPhase.eFault; // 迁故障相 / migrate to the fault phase
END_CASE

// 段 6｜失能与故障最终否决：命令一律受故障锁存与失能否决 / segment 6, final veto by the fault latch and the enable
IF _bFault OR (NOT bEnable) THEN // 故障锁存或失能 / fault latched or disabled
    bLoadCmd := FALSE; // 撤上料命令 / withdraw the load command
    bStackCmd := FALSE; // 撤叠片命令 / withdraw the stack command
    bPressCmd := FALSE; // 撤压紧命令 / withdraw the press command
    bSealCmd := FALSE; // 撤封口命令 / withdraw the seal command
    bUnloadCmd := FALSE; // 撤下料命令 / withdraw the unload command
    _bDoneInt := FALSE; // 撤周期完成脉冲内部位 / withdraw the internal cycle done bit
END_IF
IF NOT bEnable THEN // 失能 / disabled
    _ePhase := E_DL_CcaPhase.eIdle; // 回空闲相 / return to idle
END_IF

// 段 7｜统一出口 / segment 7, unified outlet
bCycleDone := _bDoneInt; // 周期完成脉冲映射本拍值 / map the cycle done pulse for this scan
_bDoneInt := FALSE; // 映射后立即撤销，保证单拍宽度（R187 两段式）/ revoke right after mapping to keep a single-scan width
nCycleCnt := _nCycle; // 周期计数出口 / cycle count outlet
bBusy := (_ePhase <> E_DL_CcaPhase.eIdle) AND (_ePhase <> E_DL_CcaPhase.eFault); // 忙指示（挂相位状态量）/ busy indicator derived from the phase state
ePhase := _ePhase; // 相位出口单点映射 / single-point phase outlet mapping
eCause := _eFaultCause; // 成因出口：全部成因均为故障级，锁存回放（R56 简化，原信息级死变量已删）/ the cause outlet, every cause is fault grade and replayed from the latch
bError := _bFault; // 故障标志与锁存位同源 / the fault flag shares the latch source
END_FUNCTION_BLOCK

(* ---- FB_DL_ColumnDpSteadyWatch.st ---- *)
(*==============================================================================
 * 组件名称 (Component)  : FB_DL_ColumnDpSteadyWatch
 * 所属子库 (Sublibrary) : DL_Process
 * 归属目录 (Directory)  : C:\Library\DL_Process
 * 当前版本 (Version)    : 1.0.0
 * 分类/来源标签         : 功能块（FUNCTION_BLOCK）· 过程监视 · 精馏塔差压
 *                         industry-pool / distillation / steady-state-watch
 * 兼容性   (Platform)   : CODESYS 3.5 / TwinCAT 3 / 汇川 InoProShop / 施耐德
 *                         Machine Expert；仅用 Standard.library 的 TON
 * 溯源声明 (Provenance) : 道莅自研 clean-room——只借公开规范条款与工程惯例，零代码行复制。
 * 功能一句话 (Summary)  : 精馏塔压差稳态监视：稳态窗学习均值与散布，稳态建立后
 *                         按液泛/漏液双阈值预判，非稳态期间抑制判定保守输出。
 *
 * 功能描述 (Function)   : 空闲相等使能转学习；学习相按节拍采样压差并跟踪
 *                         最小/最大值，窗满时均值与散布一次导出，散布不超过
 *                         均值的稳态带百分比则宣告稳态（信息级 3005），否则
 *                         报 3007 重学习；监视相输出偏差百分比，压差越液泛
 *                         阈值报液泛风险、越漏液阈值报漏液风险。输入非有限
 *                         冻结评估（3006），非物理跳变冻结转重学习（3008）。
 * 与既有件边界 (Boundary): 前置件 FB_DL_ColumnDpCtrl 做压差调节；本件只做
 *                         稳态判定与预判，不输出操作指令，二者正交级联。
 * 码位说明 (Codes)      : 信息 16#0006_3005 稳态建立（均值与散布可用）
 *                         故障 16#0006_3006 输入非有限，评估冻结
 *                         故障 16#0006_3007 稳态窗超时未达稳态，重学习
 *                         故障 16#0006_3008 非物理跳变，判定冻结重学习
 *                         段 16#06_0_05~09 首槽信息级、次槽起故障级。
 * 依赖说明 (Depends)    : 无 DL_ 内部依赖；仅 Standard.library 的 TON。
 * 红线自检 (Redline)    : 零全局依赖 ｜ 零 VAR_EXTERNAL ｜ 零 %I/%Q ｜ 纯 IEC 标准库
 *                         浮点比较全部带 fEps 容差 ｜ NaN/Inf 精确判据拦截
 *                         ENUM 配 CASE 且 ELSE 兜底 ｜ 定时器每周期无条件刷新
 *                         全变量双语同行注释 ｜ 故障锁存回放且有可达解除路径
 * 修订历史 (Revision)   : 2026-11-18  v1.0.0  首版入库（R32 · 批 2）
 *============================================================================*)

FUNCTION_BLOCK FB_DL_ColumnDpSteadyWatch
VAR_INPUT
    bRun       : BOOL;                    // 监视使能，假则回空闲并清判定 / Enable, FALSE returns to idle
    fDpKpa     : LREAL;                   // 塔压差 [kPa] / Column differential pressure
    fBandPct   : LREAL := 5.0;            // 稳态带 [％]，散布占均值上限 / Steady band as percent of the mean
    fFloodThKpa: LREAL := 8.0;            // 液泛预判阈值 [kPa] / Flooding prejudge threshold
    fLeakThKpa : LREAL := 1.5;            // 漏液预判阈值 [kPa] / Weeping prejudge threshold
    fEps       : LREAL := 1.0E-6;         // 浮点判零容差 [实数域] / Floating zero tolerance
    tSteadyWin : TIME  := T#15M;          // 稳态窗时长 [s] / Steady window duration
    tSample    : TIME  := T#5S;           // 采样节拍 [s] / Sampling pace period
END_VAR
VAR_OUTPUT
    ePrejudge : (eNormal := 0, eFloodRisk := 1, eLeakRisk := 2);    // 预判枚举 / Prejudge enum
    bSteady   : BOOL;                   // 稳态标志，均值与散布可用时为真 / TRUE when steady stats are valid
    fMeanKpa  : LREAL;                  // 学习均值 [kPa] / Learned mean
    fSpreadKpa: LREAL;                  // 学习散布（最大减最小）[kPa] / Learned spread, max minus min
    fDevPct   : LREAL;                  // 当前偏差 [％]，相对学习均值 / Current deviation vs the mean
    bError    : BOOL;                   // 故障标志，与故障码配对 / Fault flag paired with codes
    uErrorId  : UDINT;                  // 事件码，0 表示无事件 / Event code, zero means none
END_VAR
VAR
    eState    : (eIdle := 0, eLearning := 1, eWatching := 2);   // 状态机：空闲/学习/监视 / State machine
    tonWin    : TON;    // 稳态窗定时器 [s]，每拍无条件刷新 / Steady window timer
    tonPace   : TON;    // 采样节拍定时器 [s]，每拍无条件刷新 / Sampling pace timer
    bSigOk    : BOOL;   // 输入有效标志 / Input validity flag
    fSumKpa   : LREAL;  // 学习相累加和 [kPa] / Learning-phase sum
    nSamples  : UDINT;  // 有效样本数 [个] / Valid sample count
    fMinKpa   : LREAL;  // 窗内最小值 [kPa] / Window minimum
    fMaxKpa   : LREAL;  // 窗内最大值 [kPa] / Window maximum
    fDpLast   : LREAL;  // 上拍压差快照 [kPa] / Previous pressure snapshot
    bHavePrev : BOOL;   // 快照有效标志 / Snapshot availability flag
    uCodeLatch: UDINT;  // 故障锁存码 [码]，故障相回放 / Latched fault code
    uInfoCode : UDINT;  // 信息级单拍码 [码] / One-shot info code
END_VAR
VAR CONSTANT
    DL_CDS_MINSAMP : INT   := 8;        // 稳态窗最小样本数 [个] / Minimum window samples
    DL_CDS_JUMP    : LREAL := 5.0;      // 单拍非物理跳变门限 [kPa] / Non-physical jump limit
    DL_CDS_PCT     : LREAL := 100.0;    // 百分比系数 [％] / Percent factor
END_VAR

(* 段 1｜定时器无条件周期刷新（红线 7）/ Timers refreshed unconditionally every scan *)
tonWin(IN := (eState = eLearning) AND bRun, PT := tSteadyWin);  // 稳态窗计时 / Steady window timing
tonPace(IN := bRun, PT := tSample);                             // 采样节拍计时 / Sampling pace timing

(* 段 2｜输入有效性（每拍计算，判据门控挂状态量）/ Input validity each scan *)
bSigOk := (fDpKpa = fDpKpa)                     // NaN 自反判据 / NaN reflexivity
          AND (ABS(fDpKpa) < 1.0E308)           // Inf 上限判据 / Inf limit
          AND (fDpKpa >= -fEps);                // 压差非负物理约束 / Physical non-negativity

(* 段 3｜状态机主分派（ENUM 配 CASE，ELSE 兜底）/ State dispatch with ELSE interception *)
CASE eState OF

    eIdle:
        bSteady := FALSE;               // 非稳态不出统计 / No stats before steady
        ePrejudge := eNormal;           // 默认预判 / Default prejudge
        fSumKpa := 0.0;                 // 清累加 / Clear the sum
        nSamples := 0;                  // 清计数 / Clear the count
        fMinKpa := 1.0E308;             // 最小值初值为上界 / Min seeded with the upper bound
        fMaxKpa := -1.0E308;            // 最大值初值为下界 / Max seeded with the lower bound
        bHavePrev := FALSE;             // 清快照 / Clear the snapshot
        IF bRun AND bSigOk THEN
            eState := eLearning;        // 拍 N 空闲相满足，拍 N+1 转学习 / Idle to learning next scan
        END_IF

    eLearning:
        (* 本拍行为：节拍到点采样并跟踪极值；退出条件 = 窗满 AND 样本足（双条件）
         * This scan: sample on pace tick; exit needs window done AND enough samples *)
        IF NOT bSigOk THEN
            uCodeLatch := 16#0006_3006; // 故障：输入非有限 / Fault: non-finite input
        ELSIF tonPace.Q THEN
            fSumKpa := fSumKpa + fDpKpa;    // 累加 / Accumulate
            nSamples := nSamples + 1;       // 计数 / Count
            IF fDpKpa < fMinKpa THEN
                fMinKpa := fDpKpa;          // 更新最小 / Update the minimum
            END_IF
            IF fDpKpa > fMaxKpa THEN
                fMaxKpa := fDpKpa;          // 更新最大 / Update the maximum
            END_IF
        END_IF
        IF tonWin.Q AND (nSamples >= INT_TO_UDINT(DL_CDS_MINSAMP)) THEN
            fMeanKpa   := fSumKpa / UDINT_TO_LREAL(nSamples);       // 均值导出 / Derive the mean
            fSpreadKpa := fMaxKpa - fMinKpa;                        // 散布导出 / Derive the spread
            IF fSpreadKpa <= (ABS(fMeanKpa) * fBandPct / DL_CDS_PCT) THEN
                bSteady := TRUE;            // 散布在带内，稳态成立 / Spread inside the band, steady
                uCodeLatch := 16#0000_0000; // 成功清除锁存 / Success clears the latch
                uInfoCode := 16#0006_3005;  // 信息级：稳态建立（单拍）/ Info: steady built, one shot
                eState := eWatching;        // 拍 N+1 转监视 / To watching next scan
            ELSE
                uCodeLatch := 16#0006_3007; // 故障：窗满未达稳态 / Fault: window done, not steady
                fSumKpa := 0.0;             // 清累加重学 / Clear for relearning
                nSamples := 0;              // 清计数 / Clear the count
                fMinKpa := 1.0E308;         // 重置极值 / Reseed the extremes
                fMaxKpa := -1.0E308;
            END_IF
        ELSIF tonWin.Q THEN
            uCodeLatch := 16#0006_3007;     // 故障：窗满样本不足 / Fault: window done, too few samples
            fSumKpa := 0.0;                 // 清累加重学 / Clear for relearning
            nSamples := 0;                  // 清计数 / Clear the count
            fMinKpa := 1.0E308;             // 重置极值 / Reseed the extremes
            fMaxKpa := -1.0E308;
        END_IF

    eWatching:
        IF NOT bSigOk THEN
            uCodeLatch := 16#0006_3006;     // 故障：输入非有限，判定冻结 / Fault: non-finite, frozen
        ELSIF ABS(fMeanKpa) < fEps THEN
            uCodeLatch := 16#0006_3008;     // 故障：基线异常，转重学习 / Fault: bad baseline, relearn
            bSteady := FALSE;               // 撤稳态标志 / Withdraw steady
            fSumKpa := 0.0;                 // 清累加 / Clear the sum
            nSamples := 0;                  // 清计数 / Clear the count
            fMinKpa := 1.0E308;             // 重置极值 / Reseed
            fMaxKpa := -1.0E308;
            eState := eLearning;            // 拍 N+1 转学习 / To learning next scan
        ELSE
            (* 非物理跳变闸：单拍超限说明取压管路异常 / Jump gate: sensing line trouble *)
            IF bHavePrev AND (ABS(fDpKpa - fDpLast) > DL_CDS_JUMP) THEN
                uCodeLatch := 16#0006_3008; // 故障：非物理跳变 / Fault: non-physical jump
                bSteady := FALSE;           // 撤稳态标志 / Withdraw steady
                fSumKpa := 0.0;             // 清累加 / Clear the sum
                nSamples := 0;              // 清计数 / Clear the count
                fMinKpa := 1.0E308;         // 重置极值 / Reseed
                fMaxKpa := -1.0E308;
                eState := eLearning;        // 拍 N+1 转学习 / To learning next scan
            ELSE
                fDevPct := (fDpKpa - fMeanKpa) / fMeanKpa * DL_CDS_PCT;     // 偏差百分比导出 / Deviation percent
                IF fDpKpa >= fFloodThKpa THEN
                    ePrejudge := eFloodRisk;    // 越液泛阈值：液泛风险 / Over flood threshold
                ELSIF fDpKpa <= fLeakThKpa THEN
                    ePrejudge := eLeakRisk;     // 越漏液阈值：漏液风险 / Under leak threshold
                ELSE
                    ePrejudge := eNormal;       // 带内正常 / Normal inside the band
                END_IF
            END_IF
        END_IF

ELSE
    eState := eIdle;                    // 非法状态拦截回空闲 / Illegal state intercepted to idle
    uCodeLatch := 16#0006_3006;         // 故障：状态越界 / Fault: state out of range
END_CASE

(* 段 4｜快照与出口装配 / Snapshot and exit assembly *)
fDpLast := fDpKpa;                      // 更新快照供下拍跳变判据 / Update the snapshot
bHavePrev := bSigOk;                    // 快照有效随数据有效 / Snapshot valid with the data
IF NOT bRun THEN
    uCodeLatch := 16#0000_0000;         // 撤使能清故障（可达解除路径）/ Run drop clears faults
END_IF
bError := (uCodeLatch <> 16#0000_0000); // 故障锁存回放 / Latched fault replay
IF uCodeLatch <> 16#0000_0000 THEN
    uErrorId := uCodeLatch;             // 故障码优先回放 / Fault code replayed first
    uInfoCode := 16#0000_0000;          // 故障压过信息码 / Fault overrides info
ELSE
    uErrorId := uInfoCode;              // 无故障时放信息码 / Info code when no fault
    uInfoCode := 16#0000_0000;          // 信息码单拍清零 / Info code cleared next scan
END_IF
END_FUNCTION_BLOCK

(* ---- FB_DL_CompressorFleetStaging.st ---- *)
(*==============================================================================
 * 组件名称 (Component)  : FB_DL_CompressorFleetStaging
 * 所属子库 (Sublibrary) : DL_Process
 * 归属目录 (Directory)  : C:\Library\DL_Process
 * 当前版本 (Version)    : 1.0.1
 * 分类/来源标签         : 功能块（FUNCTION_BLOCK）· 公用工程 · 空压机群站编排
 *                         industry-pool / compressed-air / fleet-staging
 * 兼容性   (Platform)   : CODESYS 3.5 / TwinCAT 3 / 汇川 InoProShop / 施耐德
 *                         Machine Expert；仅用 Standard.library 的 TON
 * 溯源声明 (Provenance) : 道莅自研 clean-room——只借公开规范条款与工程惯例，零代码行复制。
 * 功能一句话 (Summary)  : 空压机群站加卸载编排：母管压力带定目标台数（TRUNC
 *                         进位点），错峰单台步进启停，最短运行/停止轮值防浪涌。
 *
 * 功能描述 (Function)   : 目标台数 = TRUNC((上限压力 − 母管压力) ÷ 压力带宽
 *                         × 总台数)，余量按 0.5 进位（R149 两式：先 TRUNC
 *                         再按余量进位，不写 TRUNC+1），结果钳到 0..总台数；
 *                         台数调整每错峰窗最多一台（防同时启停浪涌）；起台
 *                         轮值指针循环选机，停台优先运行时间最短者；单台
 *                         最短运行/最短停止时间由独立 TON 实例守护。
 * 与既有件边界 (Boundary): 本件只出各台加载指令，不出调节阀/变频指令；
 *                         压力闭环归调节件，本件是台数编排层。
 * 码位说明 (Codes)      : 信息 16#0006_3014 台数调整步进执行（单台错峰）
 *                         故障 16#0006_3015 压力带域外（高低倒置或带宽近零）——本拍重算，非锁存
 *                         故障 16#0006_3016 台数域外（小于 1 或大于 8）——本拍重算，非锁存
 *                         故障 16#0006_3017 压力输入非有限，编排冻结——锁存，bSigOk 恢复沿清码
 *                         段 16#06_0_14~18 首槽信息级、次槽起故障级。
 * 依赖说明 (Depends)    : 无 DL_ 内部依赖；仅 Standard.library 的 TON / ABS。
 * 红线自检 (Redline)    : 零全局依赖 ｜ 零 VAR_EXTERNAL ｜ 零 %I/%Q（台阵引脚）
 *                         除法前强制判零（带宽容差闸）｜ NaN/Inf 精确判据
 *                         ENUM 配 CASE 且 ELSE 兜底 ｜ TON 用 ARRAY 各台独立
 *                         实例且每周期无条件刷新 ｜ 全变量双语同行注释
 * 修订历史 (Revision)   : 2026-11-18  v1.0.0  首版入库（R32 · 批 3）
 *                        2026-11-18  v1.0.1  R33 返修：错峰窗自复位振荡；3015/3016 改本拍重算非锁存；3017 加恢复沿清码
 *============================================================================*)

FUNCTION_BLOCK FB_DL_CompressorFleetStaging
VAR_INPUT
    bRun        : BOOL;                     // 编排使能，假则全卸载清指针 / Enable, FALSE unloads all
    fHeaderKpa  : LREAL;                    // 母管压力 [kPa] / Header pressure
    fBandLowKpa : LREAL := 620.0;           // 压力带下限 [kPa]，低于则加台 / Band lower limit
    fBandHighKpa: LREAL := 700.0;           // 压力带上限 [kPa]，高于则减台 / Band upper limit
    nUnitsMax   : INT;                      // 可用台数 [台]，域 1 到 8 / Available units, 1 to 8
    tMinRunS    : TIME  := T#120S;          // 单台最短运行时间 [s] / Minimum run time per unit
    tMinStopS   : TIME  := T#180S;          // 单台最短停止时间 [s] / Minimum stop time per unit
    tStaggerS   : TIME  := T#30S;           // 错峰窗时长 [s]，窗内最多一台启停 / Stagger window
    fEps        : LREAL := 1.0E-6;          // 浮点判零容差 [实数域] / Floating zero tolerance
END_VAR
VAR_OUTPUT
    aStaged : ARRAY[1..8] OF BOOL;      // 各台加载指令 [引脚]，1 到 8 台 / Per-unit load commands
    nStaged : INT;                      // 当前加载台数 [台] / Currently staged count
    bError  : BOOL;                     // 故障标志，与故障码配对 / Fault flag paired with codes
    uErrorId: UDINT;                    // 事件码，0 表示无事件 / Event code, zero means none
END_VAR
VAR
    _eState    : (eStIdle := 0, eStRegulating := 1);    // 状态机：空闲/调节 / State machine
    tonStagger : TON;           // 错峰窗定时器 [s]，每拍无条件刷新 / Stagger window timer
    aTonRun    : ARRAY[1..8] OF TON;    // 各台最短运行计时（R158 独立实例）/ Per-unit run timers
    aTonStop   : ARRAY[1..8] OF TON;    // 各台最短停止计时（R158 独立实例）/ Per-unit stop timers
    bSigOk     : BOOL;          // 压力输入有效标志 / Pressure validity flag
    bBandOk    : BOOL;          // 压力带域有效标志 / Band validity flag
    iTarget    : INT;           // 目标台数 [台] / Target count
    fNeed      : LREAL;         // 台数需求比例值 [比值] / Count demand as a ratio
    fFrac      : LREAL;         // TRUNC 后余量 [比值]，进位判据 / Remainder for the carry
    fBandW     : LREAL;         // 压力带宽 [kPa] / Band width
    nRotPtr    : INT;           // 起台轮值指针 [索引]，1 到 nUnitsMax 循环 / Rotation pointer
    nI         : INT;           // 台循环下标 [索引] / Unit loop index
    uCodeLatch : UDINT;         // 故障锁存码 [码] / Latched fault code
    uInfoCode  : UDINT;         // 信息级单拍码 [码] / One-shot info code
    uLevelCode : UDINT;         // 本拍重算级故障码，非锁存（R33 返修）/ Recomputed per-scan fault code
    bSigOkPrev : BOOL;          // 上拍压力有效快照，恢复沿判据 / Previous validity snapshot
END_VAR
VAR CONSTANT
    DL_CFS_NMAX  : INT   := 8;          // 台数上限 [台]，与数组声明一致 / Unit cap, matches the array
    DL_CFS_HALF  : LREAL := 0.5;        // 进位余量阈值 [比值] / Carry remainder threshold
END_VAR

(* 段 1｜定时器无条件刷新（红线 7）：错峰窗与各台运行/停止计时全部每拍触发
 *      Timers refreshed unconditionally: stagger window plus per-unit arrays *)
tonStagger(IN := NOT tonStagger.Q, PT := tStaggerS);    // 错峰窗自复位振荡（R33 返修）/ Self-reset oscillating window
FOR nI := 1 TO DL_CFS_NMAX DO
    aTonRun[nI](IN := aStaged[nI], PT := tMinRunS); // 运行计时随加载 / Run timing with load
    aTonStop[nI](IN := NOT aStaged[nI], PT := tMinStopS);   // 停止计时随卸载 / Stop timing with unload
END_FOR

(* 段 2｜输入有效性与压力带域闸（本拍重算级：条件消失即清，非锁存）/ Validity and band gate, recomputed *)
uLevelCode := 16#0000_0000;                 // 每拍先清，条件不满足再置（可达清零）/ Clear each scan
bSigOk := (fHeaderKpa = fHeaderKpa)                 // NaN 自反判据 / NaN reflexivity
          AND (ABS(fHeaderKpa) < 1.0E308);          // Inf 上限判据 / Inf limit
bBandOk := ((fBandHighKpa - fBandLowKpa) > fEps)    // 带宽必须为正 / Band width positive
           AND (nUnitsMax >= 1) AND (nUnitsMax <= DL_CFS_NMAX);  // 台数域约束 / Count domain
IF NOT bBandOk THEN
    uLevelCode := 16#0006_3015;         // 本拍重算：压力带域外 / Recomputed: band out of domain
    IF (nUnitsMax < 1) OR (nUnitsMax > DL_CFS_NMAX) THEN
        uLevelCode := 16#0006_3016;     // 本拍重算：台数域外便于排查 / Recomputed: count out of domain
    END_IF
END_IF

(* 段 3｜状态机主分派（ENUM 配 CASE，ELSE 兜底）/ State dispatch with ELSE interception *)
CASE _eState OF

    eStIdle:
        (* 本拍行为：全卸载；使能与域闸俱备拍 N+1 转调节 / Unload all; arm when valid *)
        FOR nI := 1 TO DL_CFS_NMAX DO
            aStaged[nI] := FALSE;       // 全卸载 / Unload all
        END_FOR
        nStaged := 0;                   // 台数清零 / Clear the count
        nRotPtr := 1;                   // 轮值指针复位 / Reset the pointer
        IF bRun AND bSigOk AND bBandOk THEN
            _eState := eStRegulating;   // 拍 N 空闲相满足，拍 N+1 转调节 / To regulating next scan
        END_IF

    eStRegulating:
        (* 本拍行为：算目标台数，错峰窗内最多调一台 / Compute the target, one unit per window *)
        IF NOT bRun THEN
            _eState := eStIdle;         // 拍 N+1 回空闲卸载 / Back to idle next scan
        ELSIF NOT bSigOk THEN
            uCodeLatch := 16#0006_3017; // 故障级：压力非有限，保持现状 / Fault: non-finite, hold
        ELSIF NOT bBandOk THEN
            (* 域闸已在段 2 报码，此处保守保持现状不调台 / Band gate holds the current staging *)
        ELSE
            fBandW := fBandHighKpa - fBandLowKpa;                       // 带宽导出 / Band width
            fNeed  := (fBandHighKpa - fHeaderKpa) / fBandW * UDINT_TO_LREAL(INT_TO_UDINT(nUnitsMax));   // 需求比例 / Demand ratio
            IF fNeed < 0.0 THEN
                fNeed := 0.0;           // 超上限压力：需求钳零 / Over-high pressure: clamp to zero
            ELSIF fNeed > UDINT_TO_LREAL(INT_TO_UDINT(nUnitsMax)) THEN
                fNeed := UDINT_TO_LREAL(INT_TO_UDINT(nUnitsMax));   // 超下限压力：需求钳满 / Over-low: clamp to full
            END_IF
            iTarget := LREAL_TO_DINT(TRUNC(fNeed));     // R149 两式：先 TRUNC / TRUNC first
            fFrac := fNeed - TRUNC(fNeed);              // 余量导出 / Remainder
            IF fFrac >= DL_CFS_HALF THEN
                iTarget := iTarget + 1;                 // 按余量进位（不是 TRUNC+1）/ Carry by remainder
            END_IF
            IF iTarget > nUnitsMax THEN
                iTarget := nUnitsMax;                   // 钳满 / Clamp full
            ELSIF iTarget < 0 THEN
                iTarget := 0;                           // 钳零 / Clamp zero
            END_IF
            (* 错峰步进：窗满且目标与现状不等时调一台，方向由目标决定
             * One unit per stagger window, direction from the target *)
            IF tonStagger.Q AND (iTarget <> nStaged) THEN
                IF iTarget > nStaged THEN
                    (* 加台：轮值指针循环找一台未加载且停止计时已满的机
                     * Stage up: rotate to a unit unloaded with its stop time served *)
                    FOR nI := 0 TO (DL_CFS_NMAX - 1) DO
                        nRotPtr := (nRotPtr MOD DL_CFS_NMAX) + 1;       // 指针循环推进 / Rotate the pointer
                        IF (NOT aStaged[nRotPtr]) AND (nRotPtr <= nUnitsMax) AND aTonStop[nRotPtr].Q THEN
                            aStaged[nRotPtr] := TRUE;   // 加载该台 / Load the unit
                            uInfoCode := 16#0006_3014;  // 信息级：步进执行 / Info: step executed
                            EXIT;                       // 单台即止 / One unit only
                        END_IF
                    END_FOR
                ELSE
                    (* 减台：找一台已加载且运行计时已满的机（最短运行守护）
                     * Stage down: a loaded unit with its run time served *)
                    FOR nI := 1 TO nUnitsMax DO
                        IF aStaged[nI] AND aTonRun[nI].Q THEN
                            aStaged[nI] := FALSE;       // 卸载该台 / Unload the unit
                            uInfoCode := 16#0006_3014;  // 信息级：步进执行 / Info: step executed
                            EXIT;                       // 单台即止 / One unit only
                        END_IF
                    END_FOR
                END_IF
                nStaged := 0;               // 台数重算 / Recount
                FOR nI := 1 TO DL_CFS_NMAX DO
                    IF aStaged[nI] THEN
                        nStaged := nStaged + 1;     // 累加实载台数 / Count the loaded units
                    END_IF
                END_FOR
            END_IF
        END_IF

ELSE
    _eState := eStIdle;                 // 非法状态拦截回空闲 / Illegal state to idle
    uCodeLatch := 16#0006_3015;         // 故障：状态越界 / Fault: state out of range
END_CASE

(* 段 4｜出口装配：3017 锁存带 bSigOk 恢复沿清码；3015/3016 本拍重算直出 / Exit assembly *)
IF (uCodeLatch = 16#0006_3017) AND bSigOk AND (NOT bSigOkPrev) THEN
    uCodeLatch := 16#0000_0000;         // 压力恢复上升沿清 3017（可达解除）/ Recovery edge clears 3017
END_IF
bSigOkPrev := bSigOk;                   // 有效标志快照 / Validity snapshot
IF NOT bRun THEN
    uCodeLatch := 16#0000_0000;         // 撤使能清故障（可达解除）/ Run drop clears faults
END_IF
IF uCodeLatch <> 16#0000_0000 THEN
    bError := TRUE;                     // 锁存故障在报 / Latched fault active
    uErrorId := uCodeLatch;             // 故障码优先 / Fault first
ELSIF uLevelCode <> 16#0000_0000 THEN
    bError := TRUE;                     // 本拍重算级故障在报 / Recomputed fault active
    uErrorId := uLevelCode;             // 域闸码本拍直出 / Band gate code this scan
ELSE
    bError := FALSE;                    // 无故障 / No fault
    uErrorId := uInfoCode;              // 信息码单拍 / Info one shot
END_IF
uInfoCode := 16#0000_0000;              // 信息码单拍消费 / Consume info code
END_FUNCTION_BLOCK
